(* IEC 61131-3 sources: daoli-st-library/DL_MathData (part 11) *)

(* ---- FC_DL_CubicBezierEval.st ---- *)
(*==============================================================================
 * 组件名称 (Component)  : FC_DL_CubicBezierEval
 * 所属子库 (Sublibrary) : DL_MathData
 * 当前版本 (Version)    : 1.0.0
 * 兼容性   (Platform)   : CODESYS 3.5+ / TwinCAT 3 / 汇川 InoProShop / 施耐德 Machine Expert
 *                         仅依赖 Standard.library 与 LREAL 四则运算，零厂商私有库
 * 功能描述 (Function)   : 一维标量三次贝塞尔曲线求值。给定四个控制点 P0~P3 与参数 t，
 *                         按 De Casteljau 递推（三级线性插值）求点值 fValue，并给出对 t 的
 *                         一阶导数 fTangent。选择 De Casteljau 而非多项式展开的理由：三次
 *                         Bernstein 展开在 t 接近 0/1 时会出现大系数相消（P0 与 P1 量级接近时
 *                         有效位丢失），De Casteljau 每级只做凸组合，数值稳定且中间量有界。
 * 分工声明 (Scope)      : 本件是**参数曲线求值**（已知控制点，求任意 t 处点与切线）；
 *                         `FC_DL_CubicSplineInterp` 是**数据点插值**（已知离散样本点，构造
 *                         分段三次样条后插值）。二者数学对象不同（Bernstein 基 vs 三次样条基），
 *                         不可互换调用：把本件当插值用会得到穿过控制包络的曲线而非过样本点曲线。
 * 接口     (Interface)  : 输入 fP0 / fP1 / fP2 / fP3 四个控制点标量值、fT 曲线参数（域 [0,1]，
 *                         越域钳制）；输出 fValue 点值、fTangent 一阶导数值、bClamped 参数
 *                         越域钳制标记、uErrorId 事件码；返回值 BOOL = TRUE 表示本次结果有效。
 * 边界     (Boundary)   : ① 参数越域（fT < 0 或 fT > 1）钳到端点并置 bClamped，不报错（钳制
 *                         是可预期的调用方行为，非故障）；
 *                         ② 任一输入非有限（NaN / ±Inf）→ 输出 0、置故障码、返回 FALSE，
 *                         绝不向下游传播 NaN（下游联锁会把 NaN 比较结果全判 FALSE 而静默失效）；
 *                         ③ 结果非有限复检兜底（防御纵深，正常域内不可能触发）；
 *                         ④ 纯函数零状态，无 TON / 边沿实例（R6 / R7 本件标注 N/A：无顺序状态机，
 *                         无实例调用，非法状态不可能出现）；
 *                         ⑤ 零全局耦合（无 GVL / 无物理地址）。
 * 判等例外 (Exception)  : 本件非有限判定使用 `x <> x`（NaN 自反）与 `(x-x) <> (x-x)`（Inf 差值
 *                         自减），此为**浮点判等禁令的唯一例外**（R79 / 机检 G6 白名单），
 *                         不得据此推断本件允许对量值使用 `=` / `<>`：量值比较在本件中不存在。
 * 码表     (Codes)      : 16#0001_03ED 故障级：贝塞尔求值故障（输入非有限 / 输出非有限复检失败），
 *                         本件单码，不细分（纯函数无归因成员，原因由入参侧唯一确定）。
 *                         16#0001_04B0 信息级：本次求值正常完成（供上层区分「未调用」与「调用成功」）。
 *                         加码反证（R90）：正常完成与「参数被钳制」在 fValue / fTangent 上不可区分
 *                         （钳制后 t 落到端点，结果与恰好传入端点值完全一致），故须以一码留痕；
 *                         钳制本身另有 bClamped 布尔出口，不再单立钳制码。
 *                         码段说明：0001 段故障子带 03xx / 信息子带 04xx，本件取 03ED / 04B0
 *                         （源码实扫该两槽为空，续接同子带已用最大值，未回填碎片孔洞）。
 * 开源溯源 (Origin)     : 道莅自研 clean-room（参考 Bernstein 基与 De Casteljau 公开算法定义，
 *                         零代码行复制；t2-1-lgf 数学子族）
 * 修订历史 (Revision)   : 2026-11-19  v1.0.0  R45 首版（批次 1 · 序号 4）
 *==============================================================================*)

FUNCTION FC_DL_CubicBezierEval : BOOL
VAR_INPUT
    fP0 : LREAL := 0.0;      // 控制点 P0 标量值（曲线起点），须有限 [工程单位] / Control point P0, curve start, must be finite
    fP1 : LREAL := 0.0;      // 控制点 P1 标量值（起点切线方向控制），须有限 [工程单位] / Control point P1, start tangent control
    fP2 : LREAL := 0.0;      // 控制点 P2 标量值（终点切线方向控制），须有限 [工程单位] / Control point P2, end tangent control
    fP3 : LREAL := 0.0;      // 控制点 P3 标量值（曲线终点），须有限 [工程单位] / Control point P3, curve end
    fT  : LREAL := 0.0;      // 曲线参数，有效域 0.0 ~ 1.0（越域钳制） [-] / Curve parameter, domain 0.0..1.0, out-of-range clamped
END_VAR
VAR_OUTPUT
    fValue   : LREAL;        // 曲线点值 B(t) [工程单位] / Curve point value B(t)
    fTangent : LREAL;        // 一阶导数 dB/dt（对 t 求导，非对弧长） [工程单位/参数] / First derivative dB/dt w.r.t. t
    bClamped : BOOL;         // 参数越域钳制标记 [-] / Parameter clamp flag
    uErrorId : UDINT;        // 事件码，0 = 无事件 / Event code, 0 = no event
END_VAR
VAR
    fTs      : LREAL;        // 钳制后的参数 t [-] / Clamped parameter t
    fOmT     : LREAL;        // 补参数 (1 - t) [-] / Complement parameter (1 - t)
    fQ0      : LREAL;        // 一级插值节点 Q0 [工程单位] / Level-1 node Q0
    fQ1      : LREAL;        // 一级插值节点 Q1 [工程单位] / Level-1 node Q1
    fQ2      : LREAL;        // 一级插值节点 Q2 [工程单位] / Level-1 node Q2
    fR0      : LREAL;        // 二级插值节点 R0 [工程单位] / Level-2 node R0
    fR1      : LREAL;        // 二级插值节点 R1 [工程单位] / Level-2 node R1
    fDiff01  : LREAL;        // 控制点差 P1 - P0 [工程单位] / Control point difference P1 - P0
    fDiff12  : LREAL;        // 控制点差 P2 - P1 [工程单位] / Control point difference P2 - P1
    fDiff23  : LREAL;        // 控制点差 P3 - P2 [工程单位] / Control point difference P3 - P2
    bNonFin  : BOOL;         // 输入非有限判定结果 [-] / Non-finite input verdict
END_VAR
VAR CONSTANT
    DL_BEZ_ORDER : LREAL := 3.0;   // 三次曲线阶数乘子（导数系数），编译期常量 [-] / Cubic order multiplier for derivative, compile-time constant
END_VAR

(* —— 段 1：返回值与输出预置（任何早退路径都不留脏值） —— *)
FC_DL_CubicBezierEval := FALSE;      // 返回值预置无效 / Preset return value invalid
fValue   := 0.0;                     // 点值预置 0，故障相即安全侧 / Point value preset 0, safe side in fault
fTangent := 0.0;                     // 切线预置 0 / Tangent preset 0
bClamped := FALSE;                   // 钳制标记预置 FALSE / Clamp flag preset FALSE
uErrorId := 16#0000_0000;            // 事件码预置无事件 / Event code preset none

(* —— 段 2：域闸（先判后算，禁算完再兜） —— *)
bNonFin := (fP0 <> fP0) OR (fP1 <> fP1) OR (fP2 <> fP2) OR (fP3 <> fP3) OR (fT <> fT)          // NaN 自反判（判等禁令唯一例外） / NaN self-reflexive test
        OR ((fP0 - fP0) <> (fP0 - fP0)) OR ((fP1 - fP1) <> (fP1 - fP1))                        // P1 差值自减判 Inf / Inf test on P1 via self-subtraction
        OR ((fP2 - fP2) <> (fP2 - fP2)) OR ((fP3 - fP3) <> (fP3 - fP3))                        // P2 / P3 差值自减判 Inf / Inf test on P2 and P3
        OR ((fT - fT) <> (fT - fT));                                                            // 参数差值自减判 Inf / Inf test on the parameter
IF bNonFin THEN
    uErrorId := 16#0001_03ED;        // 故障级：输入非有限，输出保持 0 / Fault-level: non-finite input, outputs stay zero
    RETURN;                          // 不抛异常，直接带码返回 / Return with code, no exception
END_IF

(* —— 段 3：参数钳制（越域钳到 [0,1] 并置标记） —— *)
IF fT < 0.0 THEN
    fTs := 0.0;                      // 下界钳制 / Clamp to lower bound
    bClamped := TRUE;                // 置钳制标记 / Set clamp flag
ELSIF fT > 1.0 THEN
    fTs := 1.0;                      // 上界钳制 / Clamp to upper bound
    bClamped := TRUE;                // 置钳制标记 / Set clamp flag
ELSE
    fTs := fT;                       // 域内直通 / Pass through inside domain
END_IF
fOmT := 1.0 - fTs;                   // 补参数 (1 - t) / Complement parameter

(* —— 段 4：De Casteljau 三级递推（委托内核，凸组合有界） —— *)
fQ0 := fOmT * fP0 + fTs * fP1;       // 一级插值 Q0 / Level-1 interpolation Q0
fQ1 := fOmT * fP1 + fTs * fP2;       // 一级插值 Q1 / Level-1 interpolation Q1
fQ2 := fOmT * fP2 + fTs * fP3;       // 一级插值 Q2 / Level-1 interpolation Q2
fR0 := fOmT * fQ0 + fTs * fQ1;       // 二级插值 R0 / Level-2 interpolation R0
fR1 := fOmT * fQ1 + fTs * fQ2;       // 二级插值 R1 / Level-2 interpolation R1
fValue := fOmT * fR0 + fTs * fR1;    // 三级插值 = 曲线点值 / Level-3 interpolation = curve point value
fDiff01 := fP1 - fP0;                // 起点段差 / Start segment difference
fDiff12 := fP2 - fP1;                // 中段差 / Middle segment difference
fDiff23 := fP3 - fP2;                // 终点段差 / End segment difference
fTangent := DL_BEZ_ORDER * ( fOmT * fOmT * fDiff01
                           + 2.0 * fOmT * fTs * fDiff12
                           + fTs * fTs * fDiff23 );   // Bernstein 导数式 dB/dt / Bernstein derivative dB/dt

(* —— 段 5：结果非有限复检兜底（防御纵深） —— *)
IF (fValue <> fValue) OR ((fValue - fValue) <> (fValue - fValue))
   OR (fTangent <> fTangent) OR ((fTangent - fTangent) <> (fTangent - fTangent)) THEN
    fValue   := 0.0;                 // 复检失败：点值归 0 / Recheck failed: point value zeroed
    fTangent := 0.0;                 // 复检失败：切线归 0 / Recheck failed: tangent zeroed
    uErrorId := 16#0001_03ED;        // 故障级：输出非有限 / Fault-level: non-finite output
    RETURN;                          // 带码返回 / Return with code
END_IF

(* —— 段 6：正常出口 —— *)
uErrorId := 16#0001_04B0;            // 信息级：求值正常完成 / Info-level: evaluation completed
FC_DL_CubicBezierEval := TRUE;       // 返回值置有效 / Return value valid

END_FUNCTION

(* ---- FC_DL_CubicSplineInterp.st ---- *)
(*
  FC_DL_CubicSplineInterp  —  自然三次样条插值与斜率输出 / Natural cubic spline interpolation with slope output
  分类 Category : DL_MathData
  码位 Code     : 16#05_0_01
  版本 Version  : 1.0.0
  来源标签 Tag  : t2-1-lgf-math
  溯源 Source   : LGF Math 语义借鉴 · clean-room 实现，仅借分类/参数域/命名，未复制源码行
  功能 Function : 1) 自然三次样条（二阶导三对角求解，Thomas 追赶法，WHILE 带死锁计数器上限 = 节点数 + 1）；
                  2) 同时输出插值值与一阶导数（斜率），供曲线跟踪/前馈使用；
                  3) 越界不外推：钳到端点并置 bInRange := FALSE。
  边界 Boundary : ① nPointCount < 2 判无效；
                  ② 节点 X 非严格递增（含相等）拒绝求值并置码，不做静默排序；
                  ③ fQueryX 越界 → 钳到端点、bInRange := FALSE、不外推；
                  ④ 三对角主元近零（|主元| < 1E-12）判节点病态置码；
                  ⑤ 节点数超 nMaxNode 组态上限拒绝（防静态数组越界）；
                  ⑥ 节点坐标非有限（NaN/Inf）拒绝求值（FB32-7 保持槽非有限闸）。
  依赖 Depends  : 无（纯 IEC 61131-3 标准运算，零库内内核可委托；SQRT/MOD 原语未使用）

  码表 Error codes（本件格 05_0_01，子码步进 +0x10）:
    16#0005_0501 故障级：组态非法（节点数 < 2 / 节点数超 nMaxNode / 节点 X 非严格递增 / 主元近零病态 / 节点非有限）
    16#0005_0511 信息级：查询点越界已钳到端点且不外推（不置 bError）

  修订历史 Revision :
    2026-11-18  v1.0.0  R36 首版入库（W1 窗次件）
*)

FUNCTION FC_DL_CubicSplineInterp : BOOL
VAR_INPUT
    afX        : ARRAY[0..63] OF LREAL;   // 节点横坐标表，要求严格递增 [任意工程单位] / Knot abscissa table, strictly increasing
    afY        : ARRAY[0..63] OF LREAL;   // 节点纵坐标表 [任意工程单位] / Knot ordinate table
    nPointCount : UINT := 0;              // 有效节点数 [个]，域 2 ~ nMaxNode / Effective knot count, domain 2..nMaxNode
    nMaxNode   : UINT := 64;              // 组态节点上限 [个]，域 2 ~ 64（静态数组上界保护）/ Configured max knot count
    fQueryX    : LREAL := 0.0;            // 查询横坐标 [任意工程单位] / Query abscissa
END_VAR
VAR_OUTPUT
    fOutY      : LREAL;                   // 插值结果 [任意工程单位]，无效时为 0 / Interpolated ordinate, 0 when invalid
    fOutSlope  : LREAL;                   // 一阶导数（斜率）[单位/单位]，无效时为 0 / First derivative, 0 when invalid
    bInRange   : BOOL;                    // 查询点是否落在节点区间内（FALSE 表示已钳到端点）/ Query inside knot span
    bValid     : BOOL;                    // 结果有效标志 / Result valid flag
    bError     : BOOL;                    // 故障标志，与故障级码配对 / Fault flag paired with fault code
    nErrId     : UDINT;                   // 事件码，0 = 无事件 / Event code, 0 = no event
END_VAR
VAR
    nCount     : INT;                                  // 生效节点数整型副本 [个] / Integer copy of knot count
    nLast      : INT;                                  // 末节点索引（nCount - 1）[1] / Last knot index
    i          : INT;                                  // 三对角求解行索引 [1] / Tridiagonal row index
    nGuard     : INT;                                  // 追赶快照死锁计数器 [1] / Back-substitution deadlock counter
    fHiPrev    : LREAL;                                // 左邻区间宽度 x[i]-x[i-1] [单位] / Left span width
    fHiNext    : LREAL;                                // 右邻区间宽度 x[i+1]-x[i] [单位] / Right span width
    fAlpha     : LREAL;                                // 追赶法右端项 [单位] / Thomas right-hand term
    fPivot     : LREAL;                                // 主元（对角元）[单位] / Pivot of tridiagonal system
    fQuery     : LREAL;                                // 生效查询横坐标（钳定后）[单位] / Effective (clamped) query abscissa
    fH         : LREAL;                                // 命中区间宽度 [单位] / Hit span width
    fA         : LREAL;                                // 左权 (x[i+1]-q)/h [1] / Left blend weight
    fB         : LREAL;                                // 右权 (q-x[i])/h [1] / Right blend weight
    nSeg       : INT;                                   // 命中区间左端索引 [1] / Hit span left index
    bFound     : BOOL;                                  // 区间查找命中标志 / Span found flag
    bMono      : BOOL;                                  // 节点严格递增检查标志 / Strict monotonic check flag
    bBad       : BOOL;                                  // 节点非有限标志 / Non-finite knot flag
    afM        : ARRAY[0..63] OF LREAL;                // 二阶导解向量 m[i] [单位] / Second derivative solution vector
    afL        : ARRAY[0..63] OF LREAL;                // 追赶法下对角 l[i] [单位] / Thomas lower diagonal
    afMu       : ARRAY[0..63] OF LREAL;                // 追赶法消元系数 mu[i] [1] / Thomas elimination coefficient
    afZ        : ARRAY[0..63] OF LREAL;                // 追赶法变换后右端 z[i] [单位] / Thomas transformed right-hand side
END_VAR
VAR CONSTANT
    DL_NODE_MIN : UINT  := 2;               // 节点数下限 [个]，单点无法定义斜率 / Minimum knot count
    DL_NODE_MAX : UINT  := 64;              // 节点数硬上限 [个]，等于数组上界 + 1 / Hard upper bound of knots
    DL_PIVOT_EPS : LREAL := 1.0E-12;       // 主元判零容差 [1]，低于此值判病态 / Pivot zero tolerance
    DL_EPS      : LREAL := 1.0E-12;        // 通用判零容差 [1] / Generic zero tolerance
END_VAR

(* —— 段 0：返回值与输出预置安全值 —— *)
FC_DL_CubicSplineInterp := FALSE;   // 返回布尔：FALSE = 本拍无有效结果
fOutY     := 0.0;                   // 插值结果预置 0
fOutSlope := 0.0;                   // 斜率预置 0
bInRange  := FALSE;                 // 区间内标志预置 FALSE
bValid    := FALSE;                 // 有效标志预置 FALSE
bError    := FALSE;                 // 故障标志预置 FALSE
nErrId    := 0;                     // 事件码预置 0
bFound    := FALSE;                 // 区间查找标志预置 FALSE
bMono     := TRUE;                  // 单调性假定成立
bBad      := FALSE;                 // 非有限假定不成立
nCount    := UINT_TO_INT(nPointCount);  // 节点数整型副本 [个]

(* —— 段 1：组态域闸（节点数与上限，先于任何数组访问） —— *)
IF (nCount < DL_NODE_MIN) OR (nCount > DL_NODE_MAX) THEN
    nErrId := 16#0005_0501;         // 故障级：节点数越 [2, 64] 域
    bError := TRUE;                 // 故障标志置位（R45 配对）
    RETURN;                         // 域闸命中不求值
END_IF
IF (nMaxNode < DL_NODE_MIN) OR (nMaxNode > DL_NODE_MAX) THEN
    nErrId := 16#0005_0501;         // 故障级：组态上限越域
    bError := TRUE;                 // 故障标志置位（R45 配对）
    RETURN;                         // 域闸命中不求值
END_IF
IF nPointCount > nMaxNode THEN
    nErrId := 16#0005_0501;         // 故障级：实际节点数超组态上限（防越界，不静默截断）
    bError := TRUE;                 // 故障标志置位（R45 配对）
    RETURN;                         // 域闸命中不求值
END_IF
IF (fQueryX <> fQueryX) OR ((fQueryX - fQueryX) <> (fQueryX - fQueryX)) THEN
    nErrId := 16#0005_0501;         // 故障级：查询横坐标非有限
    bError := TRUE;                 // 故障标志置位（R45 配对）
    RETURN;                         // 域闸命中不求值
END_IF
nLast := nCount - 1;                // 末节点索引 [1]

(* —— 段 2：节点表体检（严格递增 + 非有限），任一不满足拒绝求值 —— *)
FOR i := 0 TO nLast DO
    IF (afX[i] <> afX[i]) OR ((afX[i] - afX[i]) <> (afX[i] - afX[i])) THEN
        bBad := TRUE;               // 节点横坐标非有限
    END_IF
    IF (afY[i] <> afY[i]) OR ((afY[i] - afY[i]) <> (afY[i] - afY[i])) THEN
        bBad := TRUE;               // 节点纵坐标非有限
    END_IF
END_FOR
IF bBad THEN
    nErrId := 16#0005_0501;         // 故障级：节点表含非有限值
    bError := TRUE;                 // 故障标志置位（R45 配对）
    RETURN;                         // 不求值
END_IF
FOR i := 1 TO nLast DO
    IF afX[i] - afX[i - 1] <= 0.0 THEN
        bMono := FALSE;             // 非严格递增（含相等与倒序）
    END_IF
END_FOR
IF NOT bMono THEN
    nErrId := 16#0005_0501;         // 故障级：节点 X 非严格递增，拒绝求值（不做静默排序）
    bError := TRUE;                 // 故障标志置位（R45 配对）
    RETURN;                         // 不求值
END_IF

(* —— 段 3：自然样条二阶导求解（Thomas 追赶法，主元近零判病态） —— *)
afM[0] := 0.0;                      // 自然边界：首端二阶导为 0
afM[nLast] := 0.0;                  // 自然边界：末端二阶导为 0
afL[0] := 1.0;                      // 追赶法初值
afMu[0] := 0.0;                     // 追赶法初值
afZ[0] := 0.0;                      // 追赶法初值
FOR i := 1 TO (nLast - 1) DO
    fHiPrev := afX[i] - afX[i - 1];                                  // 左邻区间宽度 [单位]
    fHiNext := afX[i + 1] - afX[i];                                  // 右邻区间宽度 [单位]，递增性已证明 > 0
    fAlpha := 3.0 / fHiNext * (afY[i + 1] - afY[i]) - 3.0 / fHiPrev * (afY[i] - afY[i - 1]);  // 右端项
    fPivot := 2.0 * (afX[i + 1] - afX[i - 1]) - fHiPrev * afMu[i - 1];                        // 主元
    IF ABS(fPivot) < DL_PIVOT_EPS THEN
        nErrId := 16#0005_0501;     // 故障级：三对角主元近零，节点病态
        bError := TRUE;             // 故障标志置位（R45 配对）
        RETURN;                     // 不出结论
    END_IF
    afL[i] := fPivot;                                               // 保存消元主元
    afMu[i] := fHiNext / afL[i];                                    // 消元系数（主元已证明非零）
    afZ[i] := (fAlpha - fHiPrev * afZ[i - 1]) / afL[i];             // 变换后右端
END_FOR
afM[nLast] := 0.0;                  // 自然边界复核（末端）
nGuard := 0;                        // 死锁计数器清零
i := nLast - 1;                     // 回代起点
WHILE (i >= 1) AND (nGuard <= (nCount + 1)) DO
    afM[i] := afZ[i] - afMu[i] * afM[i + 1];                        // 回代求二阶导
    i := i - 1;                                                     // 索引递减
    nGuard := nGuard + 1;                                           // 死锁计数器自增
END_WHILE
IF nGuard > (nCount + 1) THEN
    nErrId := 16#0005_0501;         // 故障级：回代未在节点数 + 1 步内收敛（结构性防御）
    bError := TRUE;                 // 故障标志置位（R45 配对）
    RETURN;                         // 不出结论
END_IF

(* —— 段 4：定位命中区间（线性查找，不外推：越界钳到端点） —— *)
fQuery := fQueryX;                  // 生效查询横坐标初值
IF fQueryX < afX[0] THEN
    fQuery := afX[0];               // 左越界钳到首端，不外推
    bInRange := FALSE;              // 标记越界
ELSIF fQueryX > afX[nLast] THEN
    fQuery := afX[nLast];           // 右越界钳到末端，不外推
    bInRange := FALSE;              // 标记越界
ELSE
    bInRange := TRUE;               // 落在节点区间内
END_IF
nSeg := 0;                          // 区间左端索引初值
FOR i := 0 TO (nLast - 1) DO
    IF (fQuery >= afX[i]) AND (fQuery <= afX[i + 1]) THEN
        nSeg := i;                  // 命中区间 [x[i], x[i+1]]
        bFound := TRUE;             // 查找命中
        EXIT;                       // 唯一区间（严格递增保证）
    END_IF
END_FOR
IF NOT bFound THEN
    nSeg := nLast - 1;              // 端点等值数值落空的兜底：取末区间
END_IF

(* —— 段 5：区间内求值与斜率（h 已证明 > 0，无除零风险） —— *)
fH := afX[nSeg + 1] - afX[nSeg];                                        // 命中区间宽度 [单位]
IF fH <= 0.0 THEN
    nErrId := 16#0005_0501;         // 故障级：命中区间宽度非正（数值退化）
    bError := TRUE;                 // 故障标志置位（R45 配对）
    RETURN;                         // 不出结论
END_IF
fA := (afX[nSeg + 1] - fQuery) / fH;                                    // 左权 [1]
fB := (fQuery - afX[nSeg]) / fH;                                        // 右权 [1]
fOutY := fA * afY[nSeg] + fB * afY[nSeg + 1]
       + ((fA * fA * fA - fA) * afM[nSeg] + (fB * fB * fB - fB) * afM[nSeg + 1]) * fH * fH / 6.0;  // 插值结果
fOutSlope := (afY[nSeg + 1] - afY[nSeg]) / fH
           - (3.0 * fA * fA - 1.0) / 6.0 * fH * afM[nSeg]
           + (3.0 * fB * fB - 1.0) / 6.0 * fH * afM[nSeg + 1];           // 一阶导数

(* —— 段 6：结果非有限复检 + 越界信息码 + 有效标志 —— *)
IF (fOutY <> fOutY) OR ((fOutY - fOutY) <> (fOutY - fOutY)) THEN
    fOutY := 0.0;                   // 非有限复检兜底
    fOutSlope := 0.0;               // 斜率同步兜底
    nErrId := 16#0005_0501;         // 故障级：插值结果非有限
    bError := TRUE;                 // 故障标志置位（R45 配对）
    RETURN;                         // 不出结论
END_IF
IF NOT bInRange THEN
    nErrId := 16#0005_0511;         // 信息级：查询点越界已钳到端点（信息级不置 bError）
END_IF
bValid := TRUE;                     // 结果有效（越界钳定亦有效，但 bInRange 已置 FALSE 提示）
FC_DL_CubicSplineInterp := TRUE;    // 返回布尔：TRUE = 本拍有可交付结果

END_FUNCTION

(* ---- FC_DL_CvdFilmStressCalc.st ---- *)
(*
  DL Factory R88 | FC_DL_CvdFilmStressCalc
  功能：Stoney 式算薄膜应力 σ=E_s·t_s²/(6(1-ν)·t_f·R)，曲率半径取绝对值、符号由曲率方向给定，超 300 MPa 提示
  开源溯源：无（clean-room 自研，依据公开工艺公式 Stoney 薄膜应力式，许可证=MIT，借鉴点=公式结构）
  规则：R1-R16 全遵守；R88 简单件标量形（纯标量入参出参，无循环体、无方法、无属性、无数组）
*)
FUNCTION FC_DL_CvdFilmStressCalc : REAL
VAR_INPUT
    fSubstModulusGPa : REAL := 200.0; // 基片双轴模量 E_s（Si(100) 约 180 GPa） [GPa] / substrate biaxial modulus [GPa]
    fSubstThkUm : REAL := 725.0; // 基片厚度 t_s [µm] / substrate thickness [um]
    fPoissonNu : REAL := 0.28; // 基片泊松比 ν（Si 约 0.28） [-] / Poisson ratio [-]
    fFilmThkUm : REAL := 1.0; // 薄膜厚度 t_f（须远小于 t_s） [µm] / film thickness [um]
    fCurvRadiusM : REAL := 10.0; // 曲率半径 R（带符号：正=上凸/张应力，负=下凹/压应力） [m] / signed radius [m]
    fLimitMPa : REAL := 300.0; // 应力绝对值报警上限 [MPa] / absolute stress alarm limit [MPa]
END_VAR
VAR_OUTPUT
    fStressMPa : REAL; // 薄膜应力 σ（正=张应力，负=压应力） [MPa] / film stress, positive is tensile [MPa]
    xOverLimit : BOOL; // TRUE=应力绝对值超过上限 [-] / TRUE when the absolute value is above the limit [-]
END_VAR
VAR
    fTsM : REAL; // 基片厚度换算为 m [m] / substrate thickness in metres [m]
    fTfM : REAL; // 薄膜厚度换算为 m（除零判据） [m] / film thickness in metres, the divisor [m]
    fDenom : REAL; // 分母 6(1-ν)·t_f·R_abs（除零判据） [m²] / denominator, the divisor [m^2]
    fMagMPa : REAL; // 应力幅值（未加符号） [MPa] / stress magnitude [MPa]
END_VAR

// 段 1｜出口预置
FC_DL_CvdFilmStressCalc := -1.0; // 哨兵返回 -1（无效） [-] / sentinel return -1, invalid [-]
fStressMPa := 0.0; // 应力预置零 [MPa] / stress preset zero [MPa]
xOverLimit := FALSE; // 超限位预置 FALSE（未判定前不报警） [-] / over-limit flag preset false [-]

// 段 2｜非有限拦截 + 域闸
IF NOT (fSubstModulusGPa > -1.0E30 AND fSubstModulusGPa < 1.0E30) OR NOT (fSubstThkUm > -1.0E30 AND fSubstThkUm < 1.0E30) OR NOT (fPoissonNu > -1.0E30 AND fPoissonNu < 1.0E30) THEN
    RETURN; // 模量/基片厚/泊松比任一非有限即拒算 [-] / any non finite input rejected [-]
END_IF
IF NOT (fFilmThkUm > -1.0E30 AND fFilmThkUm < 1.0E30) OR NOT (fCurvRadiusM > -1.0E30 AND fCurvRadiusM < 1.0E30) OR NOT (fLimitMPa > -1.0E30 AND fLimitMPa < 1.0E30) THEN
    RETURN; // 膜厚/曲率半径/上限任一非有限则判据静默失效，故先拦 [-] / these pins must be finite [-]
END_IF
IF fSubstModulusGPa <= 0.0 OR fSubstThkUm < 1.0E-9 OR fFilmThkUm < 1.0E-9 THEN
    RETURN; // 模量正域闸 + 厚度正域闸（分母因子不得为零） [GPa, µm] / positive modulus and thicknesses
END_IF
IF fPoissonNu <= -1.0 OR fPoissonNu >= 0.5 OR ABS(fCurvRadiusM) < 1.0E-9 OR fLimitMPa <= 0.0 THEN
    RETURN; // 泊松比开区间闸 (-1,0.5) + 曲率绝对值闸 + 上限正域闸 [-] / Poisson, radius and limit gates
END_IF

// 段 3｜计算（Stoney 式，长度统一换算到 m、模量换算到 Pa，末步转 MPa）
fTsM := fSubstThkUm * 1.0E-6; // µm × 1e-6 m/µm = m，基片厚换算 [m] / [um] x [m/um] = [m]
fTfM := fFilmThkUm * 1.0E-6; // µm × 1e-6 m/µm = m，膜厚换算 [m] / [um] x [m/um] = [m]
fDenom := 6.0 * (1.0 - fPoissonNu) * fTfM * ABS(fCurvRadiusM); // 无量纲 × 无量纲 × m × m = m²，分母 [m²] / [m^2]
IF fDenom < 1.0E-9 THEN
    RETURN; // 除法前分母闸：6(1-ν)t_f·R 必须大于 1E-9 才可作除数 [m²] / denominator gate [m^2]
END_IF
fMagMPa := fSubstModulusGPa * 1.0E9 * fTsM * fTsM / fDenom * 1.0E-6; // Pa × m² ÷ m² = Pa，再 ×1e-6 转 MPa [MPa] / [MPa]
IF fCurvRadiusM < 0.0 THEN
    fStressMPa := -fMagMPa; // 负曲率对应压应力（符号约定），幅值来自上式的绝对半径 [MPa] / compressive [MPa]
ELSE
    fStressMPa := fMagMPa; // 正曲率对应张应力（符号约定），幅值来自上式的绝对半径 [MPa] / tensile [MPa]
END_IF

// 段 4｜判定与饱和
IF NOT (fStressMPa > -1.0E30 AND fStressMPa < 1.0E30) THEN
    RETURN; // 结果非有限再拦一次（防溢出成 Inf） [MPa] / re-check the result for finiteness [MPa]
END_IF
xOverLimit := ABS(fStressMPa) > fLimitMPa; // 按绝对值与上限直比（张压同判） [MPa] / compare the magnitude [MPa]

// 段 5｜出口自检
IF fTfM >= fTsM THEN RETURN; END_IF // 出口自检：Stoney 式前提是薄膜远薄于基片，t_f>=t_s 时结果不可信 [m] / premiss violated
FC_DL_CvdFilmStressCalc := fStressMPa; // 返回薄膜应力（正=张，负=压） [MPa] / return the film stress [MPa]
END_FUNCTION

(* ---- FC_DL_DateAddDays.st ---- *)
(*
    FC_DL_DateAddDays —— DATE 加天数偏移
    ------------------------------------------------------------------
    分类      : DL_MathData / TimeArith
    前缀      : FC_DL_
    版本      : 1.0.0
    溯源      : IEC 61131-3 标准语义的道莅防御性实现（日期 + 天数 → 日期，可负偏移）；
                经天数路径委托平台内建 DATE_TO_DINT / DINT_TO_DATE 完成历法换算，
                本件不重实现历法内核；
                偏移钳位、溢出预判、双出口错误分级与码位 100% 自有；
                clean-room 重写，未复制任何闭源厂商源码，参考实现仅限 MIT/Apache 许可
    平台      : 纯 IEC 61131-3，CODESYS V3.5+ / TwinCAT 3 / InoProShop 通用
    作者      : 道莅代码库 · PLC编程专家（R20）
    ------------------------------------------------------------------
    功能说明  : 保质期到日子、交期推算、下次保养日（今天 + 90 天）、点检周期回推（今天 − 30 天）
                这类现场每天都在用的算术。日历加法不能靠秒数硬加：夏令时与闰秒都不参与
                工业日期的语义，天数路径才是唯一稳定口径。
                核心防御：① 统一走天数路径（先 DATE_TO_DINT，加偏移后再 DINT_TO_DATE），
                   不做 DT 秒级加减——秒级加减在跨闰日的边界上会差一天，而这一天
                   对保质期判定的意义不用解释；
                ② 溢出用减法比较预判，不用加法后回查符号位：nWork > 上限 − nBase
                   这类判据在任何整数表示下都成立，禁「先加再判是否变号」的写法
                   （带符号溢出的回绕行为在平台上并不一定有保证）；
                ③ 偏移超 ±36500 天（±100 年）先钳位并发信息级：排程里出现 ±100 年
                   必然是单位错（毫秒当秒填），钳位后可算但不静默；
                ④ 结果早于纪元或超容器域一律返回纪元日并置 bValid = FALSE，不做饱和——
                   饱和会伪造日期（把越界算成 1970-01-01），台账上看不出异常；
                ⑤ 天数上界与 FC_DL_DateToDintDays / FC_DL_DintDaysToDate 用同一常量口径，
                   三件之间不会错位。
                职责边界：日期差值归 FC_DL_DateDiffDays；闰年原子归 FC_DL_LeapYearChk；
                纯天数双向转换归 FC_DL_DateToDintDays / FC_DL_DintDaysToDate。
    编译门槛  : 主路径依赖平台内建 DATE_TO_DINT / DINT_TO_DATE（天数口径），
                三平台标准库均提供。天数口径的平台差异见 FC_DL_DateToDintDays 的
                编译门槛段与 DL_DATE_DAYS_MAX 的保守取值；若实测口径不同只调该常量，
                本件的闸门顺序与出口不变。
    错误码    : 16#0001_042A 偏移超 ±36500 天（±100 年）已钳位——信息级，值可用但偏移已被限幅
                16#0001_042B 预留禁用（信息级，不得挪用）
                16#0001_035D 结果早于纪元——故障级，返回纪元日
                16#0001_035E 结果超 DATE 容器域——故障级，返回纪元日，不做饱和
                16#0001_035F 预留禁用（故障级，不得挪用）
    码位总账  : 16#0001_042A 用 / 16#0001_042B 预留 ｜ 16#0001_035D 用 / 16#0001_035E 用 / 16#0001_035F 预留
    状态机    : R6 标注 N/A —— 本组件为纯函数无顺序状态机，无 CASE 可写，非法状态不可能出现
    采样约定  : 本件无定时器、无沿检测、无状态；单拍纯计算，结论与任务周期无关。
    修订记录  : 2026-11-16 v1.0.0 首次入库（R20）
*)
FUNCTION FC_DL_DateAddDays : DATE
VAR_INPUT
    dateIn           : DATE;                  // 基准日期 [日期]，有效域 1970-01-01 起 / base date [date], domain starts at 1970-01-01
    nDays            : DINT;                  // 天数偏移，可负 [日]，有效域 −36500~36500 / day offset, signed [day], valid domain −36500 to 36500
END_VAR
VAR_OUTPUT
    eErr             : UDINT;                 // 错误码，0=正常 / error id, 0=ok
    bError           : BOOL;                  // 故障标志，eErr 为故障级时 TRUE / error flag, TRUE on fault-level eErr
    bValid           : BOOL;                  // 返回值是否可用（故障级为 FALSE）/ return usable, FALSE on fault level
    bClamped         : BOOL;                  // 偏移超 ±36500 天已钳位 / the offset was clamped into the span limit
END_VAR
VAR CONSTANT
    DL_DAYS_SPAN_MAX : DINT := 36500;         // 正向偏移钳位，约 ±100 年 [日] / forward offset clamp, about one hundred years [day]
    DL_DAYS_SPAN_NEG_MAX : DINT := -36500;    // 负向偏移钳位 [日] / backward offset clamp [day]
    DL_DATE_DAYS_MIN : DINT := 0;             // 纪元日，天数下界 [日] / the epoch day, lower bound [day]
    DL_DATE_DAYS_MAX : DINT := 65535;         // 保守容器口径上限，无符号 16 位天数顶 [日] / conservative container top [day]
    DL_EPOCH_DATE_ZERO : DATE := DATE#1970-01-01; // 纪元起始日期，故障缺省返回 / the epoch date returned on faults
END_VAR
VAR
    nBase            : DINT;                  // 基准日期天数中间量 [日] / base date in days since the epoch [day]
    nWork            : DINT;                  // 偏移副本，钳位后参与加法 [日] / offset copy, used after the clamp [day]
    nOut             : DINT;                  // 结果天数中间量 [日] / result day count intermediate [day]
    nLimit           : DINT;                  // 可用余量的减法判据中间量 [日] / headroom intermediate used by the subtraction test [day]
END_VAR

// 段 1｜返回值与错误状态预置 / segment 1, preset return value and error status
FC_DL_DateAddDays := DL_EPOCH_DATE_ZERO;      // 故障缺省返回纪元日 / fault default returns the epoch date
eErr := 0;                                    // 预置无错误 / preset no error
bError := FALSE;                              // 预置无故障 / preset no fault
bValid := FALSE;                              // 预置不可用，通过闸门后置位 / preset invalid, set TRUE after the gates
bClamped := FALSE;                            // 预置未钳位 / preset no clamp
nWork := nDays;                               // 取入参副本，绝不改动调用方数据 / copy the input, never modifies caller data
nOut := DL_DATE_DAYS_MIN;                     // 结果中间量清零 / clear the result intermediate

// 段 2｜偏移跨度量闸：超 ±100 年先钳位并如实登记（信息级）/ segment 2, span gate with an explicit info-level clamp
IF nWork > DL_DAYS_SPAN_MAX THEN
    nWork := DL_DAYS_SPAN_MAX;                // 正向钳位至 +36500 天 [日] / clamp to plus 36500 days [day]
    bClamped := TRUE;                         // 标记已钳位 / flag the clamp
    eErr := 16#0001_042A;                     // 信息级：偏移超跨度已钳位 / info level, the offset was clamped
ELSIF nWork < DL_DAYS_SPAN_NEG_MAX THEN
    nWork := DL_DAYS_SPAN_NEG_MAX;            // 负向钳位至 −36500 天 [日] / clamp to minus 36500 days [day]
    bClamped := TRUE;                         // 标记已钳位 / flag the clamp
    eErr := 16#0001_042A;                     // 信息级：偏移超跨度已钳位 / info level, the offset was clamped
END_IF

// 段 3｜基准日期域闸：基准本身必须在容器域内 / segment 3, base date domain gate
nBase := DATE_TO_DINT(dateIn);                // 日期 → 自纪元天数 [日] / date to days since the epoch [day]
IF nBase < DL_DATE_DAYS_MIN THEN
    eErr := 16#0001_035D;                     // 故障级：基准日期早于纪元 / fault level, the base date precedes the epoch
    bError := TRUE;                           // 置故障标志 / raise the error flag
    bValid := FALSE;                          // 返回值不可用 / flag the return as unusable
    FC_DL_DateAddDays := DL_EPOCH_DATE_ZERO;  // 确定缺省值：纪元日 / deterministic default of the epoch date
    RETURN;                                   // 出口 / exit
END_IF
IF nBase > DL_DATE_DAYS_MAX THEN
    eErr := 16#0001_035E;                     // 故障级：基准日期超容器域 / fault level, the base date exceeds the container
    bError := TRUE;                           // 置故障标志 / raise the error flag
    bValid := FALSE;                          // 返回值不可用 / flag the return as unusable
    FC_DL_DateAddDays := DL_EPOCH_DATE_ZERO;  // 确定缺省值：纪元日 / deterministic default of the epoch date
    RETURN;                                   // 出口 / exit
END_IF

// 段 4｜正向溢出预判：用「上限 − 基准」做减法比较，禁先加后判变号 / segment 4, forward overflow test by subtraction
IF nWork > DL_DATE_DAYS_MIN THEN
    nLimit := DL_DATE_DAYS_MAX - nBase;       // 剩余可用天数 [日] / remaining room in days [day]
    IF nWork > nLimit THEN
        eErr := 16#0001_035E;                 // 故障级：结果将超 DATE 容器域 / fault level, the result would exceed the container
        bError := TRUE;                       // 置故障标志 / raise the error flag
        bValid := FALSE;                      // 返回值不可用 / flag the return as unusable
        FC_DL_DateAddDays := DL_EPOCH_DATE_ZERO; // 确定缺省值：纪元日，不伪造日期 / deterministic default, no fabricated date
        RETURN;                               // 出口 / exit
    END_IF
ELSIF nWork < DL_DATE_DAYS_MIN THEN
    // 段 5｜负向溢出预判：可用余额同为负数，比较方向不变 / segment 5, backward overflow test
    nLimit := DL_DATE_DAYS_MIN - nBase;       // 负向可用余额，负值 [日] / backward headroom, a negative value [day]
    IF nWork < nLimit THEN
        eErr := 16#0001_035D;                 // 故障级：结果将早于纪元 / fault level, the result would precede the epoch
        bError := TRUE;                       // 置故障标志 / raise the error flag
        bValid := FALSE;                      // 返回值不可用 / flag the return as unusable
        FC_DL_DateAddDays := DL_EPOCH_DATE_ZERO; // 确定缺省值：纪元日 / deterministic default of the epoch date
        RETURN;                               // 出口 / exit
    END_IF
END_IF

// 段 6｜主体：溢出已排除，加法与内建还原均安全 / segment 6, the addition and the built-in are safe after the gates
nOut := nBase + nWork;                        // 结果天数 [日] / result day count [day]
FC_DL_DateAddDays := DINT_TO_DATE(nOut);      // 天数 → 日期 / days back to a date

// 段 7｜发布结果 / segment 7, publish the result
bValid := TRUE;                               // 域内结果可用 / the in-domain result is usable
bError := FALSE;                              // 信息级不置故障（双保险）/ info level never raises a fault, second line of defence
END_FUNCTION

(* ---- FC_DL_DateDiffDays.st ---- *)
(*
    FC_DL_DateDiffDays —— 两 DATE 之差天数（可负）
    ------------------------------------------------------------------
    分类      : DL_MathData / TimeArith
    前缀      : FC_DL_
    版本      : 1.0.0
    溯源      : IEC 61131-3 标准语义的道莅防御性实现（两个日期之间的天数差，可负）；
                经天数路径委托平台内建 DATE_TO_DINT 完成历法换算，本件不重实现历法内核；
                负值口径、方向标志、错误分级与码位 100% 自有；
                clean-room 重写，未复制任何闭源厂商源码，参考实现仅限 MIT/Apache 许可
    平台      : 纯 IEC 61131-3，CODESYS V3.5+ / TwinCAT 3 / InoProShop 通用
    作者      : 道莅代码库 · PLC编程专家（R20）
    ------------------------------------------------------------------
    功能说明  : 保质期余量、超期天数、保养逾期天数的判定原子：给两个日期，输出「从前者到后者
                过了多少天」，后者早于前者即为负。与 FC_DL_DateAddDays 构成判定原子对。
                核心防御：① 差值一律在 DINT 域内做：两个 DATE 都在容器域内，天数差模长必小于
                   65536，DINT 承载结构性不溢出——此论证是本件不设故障出口的依据；
                ② 负值是合法业务输出（超期天数就是负的余量），绝不钳到 0、绝不用绝对值：
                   把「已超期 3 天」抹平成「今天到期」是保质期逻辑最典型的静默错；
                ③ bNegative 单独回告方向，HMI 不必自己再比一次大小；
                ④ 本件五槽中信息 1 槽使用、故障 3 槽按规格预留——域外输入在类型域上
                   不可表达（DATE 值域由类型系统保证），故不虚构不存在的故障码。
                职责边界：日期加偏移归 FC_DL_DateAddDays；日期天数化归 FC_DL_DateToDintDays；
                本件只管两日期之间的差值。
    编译门槛  : 主路径依赖平台内建 DATE_TO_DINT（天数口径），三平台标准库均提供。
                若某平台 DATE 以秒承载，则差值单位为秒而非天——此差异由 DL_DATE_DAYS_MAX
                的实测锚定统一裁定（与 FC_DL_DateToDintDays 同源），本件闸门不受影响。
    错误码    : 16#0001_042C 差值为负（dateTo 早于 dateFrom），已如实输出——信息级，值可用
                16#0001_042D 预留禁用（信息级，不得挪用）
                16#0001_0360 预留（故障级，不得挪用）
                16#0001_0361 预留禁用（故障级，不得挪用）
                16#0001_0362 预留禁用（故障级，不得挪用）
    码位总账  : 16#0001_042C 用 / 16#0001_042D 预留 ｜ 16#0001_0360 预留 / 16#0001_0361 预留 / 16#0001_0362 预留
    状态机    : R6 标注 N/A —— 本组件为纯函数无顺序状态机，无 CASE 可写，非法状态不可能出现
    采样约定  : 本件无定时器、无沿检测、无状态；单拍纯计算，结论与任务周期无关。
    修订记录  : 2026-11-16 v1.0.0 首次入库（R20）
*)
FUNCTION FC_DL_DateDiffDays : DINT
VAR_INPUT
    dateFrom         : DATE;                  // 区间起始日期 [日期] / start date of the interval [date]
    dateTo           : DATE;                  // 区间结束日期 [日期]，早于起点即差值为负 / end date of the interval [date], earlier than the start yields a negative difference
END_VAR
VAR_OUTPUT
    eErr             : UDINT;                 // 错误码，0=正常 / error id, 0=ok
    bError           : BOOL;                  // 故障标志，本件无故障级出口，恒为 FALSE / error flag, always FALSE here as no fault exit exists
    bValid           : BOOL;                  // 返回值是否可用（本件恒为 TRUE）/ return usable, always TRUE here
    bNegative        : BOOL;                  // 差值为负（dateTo 早于 dateFrom）/ the difference is negative
END_VAR
VAR CONSTANT
    DL_DINT_ZERO     : DINT := 0;             // 有符号零常量，避免裸字面量 [日] / signed zero constant [day]
END_VAR
VAR
    nFrom            : DINT;                  // 起始日期天数 [日] / start date in days [day]
    nTo              : DINT;                  // 结束日期天数 [日] / end date in days [day]
    nDiff            : DINT;                  // 差值中间量，可负 [日] / difference intermediate, possibly negative [day]
END_VAR

// 段 1｜返回值与错误状态预置 / segment 1, preset return value and error status
FC_DL_DateDiffDays := DL_DINT_ZERO;           // 缺省返回 0 天 [日] / default returns zero days [day]
eErr := 0;                                    // 预置无错误 / preset no error
bError := FALSE;                              // 本件无故障级出口，恒 FALSE / no fault exit exists, always FALSE
bValid := FALSE;                              // 预置不可用，末段置位 / preset invalid, set TRUE in the last stage
bNegative := FALSE;                           // 预置非负差 / preset a non-negative difference
nDiff := DL_DINT_ZERO;                        // 中间量清零 / clear the intermediate

// 段 2｜取值：两日期各做一次显式标准转换 / segment 2, both dates are converted explicitly
nFrom := DATE_TO_DINT(dateFrom);              // 起始日期天数 [日] / start date in days [day]
nTo := DATE_TO_DINT(dateTo);                  // 结束日期天数 [日] / end date in days [day]

// 段 3｜求差：模长必小于 65536，DINT 承载结构性不溢出 / segment 3, the difference cannot overflow DINT
nDiff := nTo - nFrom;                         // 有符号天数差 [日] / signed difference in days [day]

// 段 4｜负值如实输出（超期余量语义，绝不抹平）/ segment 4, negative values are published as they are
IF nDiff < DL_DINT_ZERO THEN
    bNegative := TRUE;                        // 标记差值为负 / flag the negative difference
    eErr := 16#0001_042C;                     // 信息级：差值为负，已如实输出 / info level, a negative difference was published as is
END_IF

// 段 5｜发布结果 / segment 5, publish the result
FC_DL_DateDiffDays := nDiff;                  // 输出天数差 [日] / publish the difference in days [day]
bValid := TRUE;                               // 正负差值均为合法业务输出 / both signs are legal business results
bError := FALSE;                              // 信息级不置故障（双保险）/ info level never raises a fault, second line of defence
END_FUNCTION

(* ---- FC_DL_DateToDintDays.st ---- *)
(*
    FC_DL_DateToDintDays —— DATE 到自纪元起的天数
    ------------------------------------------------------------------
    分类      : DL_MathData / Convert
    前缀      : FC_DL_
    版本      : 1.0.0
    溯源      : IEC 61131-3 标准语义的道莅防御性实现（DATE → 自 1970-01-01 起天数）；
                委托平台内建 DATE_TO_DINT 完成天数口径换算，本件不重实现历法内核；
                纪元域闸门、保守容器口径钳位、错误分级与码位 100% 自有；
                clean-room 重写，未复制任何闭源厂商源码，参考实现仅限 MIT/Apache 许可
    平台      : 纯 IEC 61131-3，CODESYS V3.5+ / TwinCAT 3 / InoProShop 通用
    作者      : 道莅代码库 · PLC编程专家（R20）
    ------------------------------------------------------------------
    功能说明  : 把日历日期折成「自 1970-01-01 起的天数」整数，供保质期、台账天数化、
                保养周期差值与数据库整型列落库使用（日期型直接落库在各家平台的位型不一致）。
                核心防御：① 早于纪元的日期在调用内建前拦下，域外调用内建可得回绕大数；
                ② 天数超保守容器口径时按容器顶钳位并发信息级，值仍可用但已注明钳位——
                   钳位事件必须可被 HMI 看见，静默钳位是本件最易漏的缺陷；
                ③ 内建返回负天数视为容器溢出（与段 2 的域门同源但不同层），单独占故障码，
                   便于区分「组态给了 1970 前日期」与「平台 DATE 位型承载异常」两类根因。
                职责边界：天数还原归 FC_DL_DintDaysToDate；带偏移的日期推算归
                FC_DL_DateAddDays；日期差值归 FC_DL_DateDiffDays。
    编译门槛  : 主路径依赖平台内建 DATE_TO_DINT（天数口径）。三平台标准库均提供该内建，
                但天数口径本身的数值锚定存在平台差异：某些平台 DATE 以秒承载、部分以天承载。
                故 DL_DATE_DAYS_MAX 取 65535（无符号 16 位天数容器上限）的保守口径，
                编码前按目标平台实测锚定；若实测口径不同，仅调本常量，闸门与出口不动。
    错误码    : 16#0001_0410 天数超保守容器口径（65535），已按容器顶钳位——信息级，值仍可用但已钳位
                16#0001_0411 预留禁用（信息级，不得挪用）
                16#0001_0336 输入日期早于纪元（1970-01-01 之前）——故障级，返回 0
                16#0001_0337 DATE 输入非法或容器溢出（内建返回负天数）——故障级，返回 0
                16#0001_0338 预留禁用（故障级，不得挪用）
    码位总账  : 16#0001_0410 用 / 16#0001_0411 预留 ｜ 16#0001_0336 用 / 16#0001_0337 用 / 16#0001_0338 预留
    状态机    : R6 标注 N/A —— 本组件为纯函数无顺序状态机，无 CASE 可写，非法状态不可能出现
    采样约定  : 本件无定时器、无沿检测、无状态；单拍纯计算，结论与任务周期无关。
    修订记录  : 2026-11-16 v1.0.0 首次入库（R20）
*)
FUNCTION FC_DL_DateToDintDays : DINT
VAR_INPUT
    dateIn           : DATE;                  // 输入日期 [日期]，有效域 1970-01-01 起 / input date [date], domain starts at 1970-01-01
END_VAR
VAR_OUTPUT
    eErr             : UDINT;                 // 错误码，0=正常 / error id, 0=ok
    bError           : BOOL;                  // 故障标志，eErr 为故障级时 TRUE / error flag, TRUE on fault-level eErr
    bValid           : BOOL;                  // 返回值是否可用（故障级为 FALSE）/ return usable, FALSE on fault level
END_VAR
VAR CONSTANT
    DL_DATE_DAYS_MIN : DINT := 0;             // 纪元日，天数下界 [日] / the epoch day, lower bound [day]
    DL_DATE_DAYS_MAX : DINT := 65535;         // 保守容器口径上限，无符号 16 位天数顶 [日] / conservative container top, unsigned 16-bit day limit [day]
    DL_EPOCH_DATE_ZERO : DATE := DATE#1970-01-01; // 纪元起始日期 / the epoch date
    DL_DINT_ZERO     : DINT := 0;             // 有符号零常量，避免裸字面量 [日] / signed zero constant [day]
END_VAR
VAR
    nDays            : DINT;                  // 自纪元起天数中间量 [日] / day count intermediate since the epoch [day]
END_VAR

// 段 1｜返回值与错误状态预置 / segment 1, preset return value and error status
FC_DL_DateToDintDays := DL_DINT_ZERO;         // 故障缺省返回 0 [日] / fault default returns zero [day]
eErr := 0;                                    // 预置无错误 / preset no error
bError := FALSE;                              // 预置无故障 / preset no fault
bValid := FALSE;                              // 预置不可用，通过闸门后置位 / preset invalid, set TRUE after the gates
nDays := DL_DINT_ZERO;                        // 中间量清零 / clear the intermediate

// 段 2｜下域闸门：早于纪元的日期先于内建拦下 / segment 2, epoch lower gate precedes the built-in call
IF dateIn < DL_EPOCH_DATE_ZERO THEN
    eErr := 16#0001_0336;                     // 故障级：输入早于纪元 / fault level, the input precedes the epoch
    bError := TRUE;                           // 置故障标志 / raise the error flag
    bValid := FALSE;                          // 返回值不可用 / flag the return as unusable
    FC_DL_DateToDintDays := DL_DINT_ZERO;     // 确定缺省值 0 / deterministic default of zero
    RETURN;                                   // 出口，不触碰内建 / exit, the built-in is never touched
END_IF

// 段 3｜主体：域内才委托平台内建（天数口径）/ segment 3, delegate the built-in only inside the domain
nDays := DATE_TO_DINT(dateIn);                // 内建换算：DATE → 自纪元天数 [日] / built-in conversion from DATE to days since the epoch [day]

// 段 4｜容器溢出闸：内建给负天数即平台 DATE 位型承载异常 / segment 4, container overflow gate
IF nDays < DL_DATE_DAYS_MIN THEN
    eErr := 16#0001_0337;                     // 故障级：DATE 非法或容器溢出 / fault level, illegal DATE or container overflow
    bError := TRUE;                           // 置故障标志 / raise the error flag
    bValid := FALSE;                          // 返回值不可用 / flag the return as unusable
    FC_DL_DateToDintDays := DL_DINT_ZERO;     // 确定缺省值 0 / deterministic default of zero
    RETURN;                                   // 出口 / exit
END_IF

// 段 5｜保守容器口径钳位（信息级，钳位事件必须可见）/ segment 5, conservative container clamp at info level
IF nDays > DL_DATE_DAYS_MAX THEN
    nDays := DL_DATE_DAYS_MAX;                // 钳位至容器顶 [日] / clamp to the container top [day]
    eErr := 16#0001_0410;                     // 信息级：超保守口径已钳位，值仍可用 / info level, clamped to the conservative top, still usable
END_IF

// 段 6｜发布结果 / segment 6, publish the result
FC_DL_DateToDintDays := nDays;                // 输出自纪元起天数 [日] / publish the days since the epoch [day]
bValid := TRUE;                               // 域内或已钳位均可用 / usable in domain or after the clamp
END_FUNCTION

(* ---- FC_DL_DateToIsoString.st ---- *)
(*
    组件名称 : FC_DL_DateToIsoString
    所属子库 : DL_MathData
    当前版本 : 1.0.1
    兼 容 性 : CODESYS V3.5+ / TwinCAT 3 / 汇川 InoProShop；仅依赖 Standard.library
    功能描述 : DATE → 'YYYY-MM-DD' 十字符定宽文本，同时把年/月/日分解结果单出口，供 MES 台账与文件名直接取用。
              取舍 ①：用 Howard Hinnant 的 civil_from_days 整数算法反算日历 —— 纯整数、无查表、无浮点、无循环，
              对任意天数一次算到位；相比「按年循环扣天数」的写法，没有循环也就没有死循环风险与扫描周期抖动。
              取舍 ②：回代自校验（days_from_civil 反算天数必须等于输入）—— 日期算法的错误往往表现为「差一天」，
              这种错在报表上极难发现，回代一次就能把「算法实现错」与「输入数据错」彻底分开；
              自校验不过就绝不输出日期。
              取舍 ③：不做平台 DATE_TO_DTL 委托 —— DTL 结构体在部分平台的字段宽度与日期语义不一致，
              且本件只需要三个整数；直接走 DATE_TO_DINT 天数口径，链路最短。
              取舍 ④：早于纪元（1970-01-01）一律判故障 —— 负数天数在部分平台 DATE 实现里是「不支持」而非「负日期」，
              与其猜，不如让调用方知道这个值不可信。
    开源溯源 : T2-1 LGF Converter 子族（只借「日期转定宽文本」这一行为定义）。civil_from_days / days_from_civil；本件为道莅 clean-room 防御性实现（仅借 LGF 分类事实/参数域/行为定义，零代码行与符号名复制）。
              为公开算法（Howard Hinnant，公有领域），本实现按整数语义重写，零代码行与注释复制；
              码位、错误分级、自校验策略 100% 自有。
    本文件内含 : FUNCTION FC_DL_DateToIsoString（单 POU，无配套类型）
    依 赖 : 无 DL_ 内部依赖；Standard.library: LEN / MID / CONCAT
    红线自检 : R1 ✓ 零全局变量与外部变量 ｜ R2 ✓ 零物理 IO 地址
              R3 ✓ 纯 IEC 61131-3 ｜ R4 ✓ 纪元闸 + 年份域闸 + 回代自校验 + 输出长度自证（全整数，无除法零风险）
              R5 ✓ 全变量中英双语同行注释 ｜ R6 N/A 纯函数无顺序状态机，无 CASE 可写
              R7 N/A 无定时器、无沿检测实例 ｜ R8 ✓ 纪元常数、闰年基数、月长基数全常量化
    错误码   : 16#0001_0450 [信息级] 输出串长异常（补零逻辑防御提示），bValid = TRUE
               16#0001_0451 [信息级] 预留禁用（不得挪用）
               16#0001_0396 [故障级] 早于纪元或年份越 1970~9999，返回 '1970-01-01'，bValid = FALSE
               16#0001_0397 [故障级] 回代自校验失败（算法自证不过），返回 '1970-01-01'，bValid = FALSE
               16#0001_0398 [故障级] 预留禁用（不得挪用）
    码位总账 : 16#0001_0450 用 / 16#0001_0451 预留 ｜ 16#0001_0396 用 / 16#0001_0397 用 / 16#0001_0398 预留
    遗留假设 : ① 【编译门槛未闭合】本件依赖「DATE_TO_DINT 返回自 1970-01-01 起的天数、纪元当日记 0」这一口径。
              CODESYS / TwinCAT 3 默认如此，InoProShop 未实测；若某平台返回秒或返回 1970-01-01 记 1，
              回代自校验会失败并置 0397（可观测，不会静默出错）。
              ② 整数除法在三平台均向零截断，本件全部操作数为非负，故截断方向不敏感 —— IEC 语义推导，未逐平台实测。
              ③ MID 参数序按 IEC 标准 MID(串, 长度, 位置)，与库内既有用法同序。
    修订历史 :
        2026-11-16  v1.0.0  首版，R21 批次 3 入库
        2026-11-16  v1.0.1  R21 终审修复（严重）：年序判据末项除数误用 DL_ERA_DAYS = 146097，
                            而 Hinnant civil_from_days 该处应为「周期内最大天序」146096。二者仅在
                            nDoe = 146096（即每个 400 年周期的最后一天 = 世纪闰日 2 月 29 日）时结果不同：
                            错值使 nYoe = 400 越出 [0, 399]，回代自校验随即失败，2000-02-29 / 2400-02-29
                            等合法日期被误判为 0397 故障并回退成 '1970-01-01'。新增常量 DL_ERA_LAST = 146096
                            并改用于该式；其余天序取值两种除数同解，故本次修复零副作用。向量已用等价脚本
                            复算：1970-01-01 / 1999-12-31 / 2000-02-29 / 2026-11-16 / 9999-12-31 全部自校验通过。
*)
FUNCTION FC_DL_DateToIsoString : STRING
VAR_INPUT
    dateIn          : DATE;   // 待格式化日期，有效域 1970-01-01 ~ 9999-12-31 / date to format, valid from 1970-01-01 to 9999-12-31
END_VAR
VAR_OUTPUT
    eErr            : UDINT;  // 错误码，0=正常；16#0001_04XX 信息级 / 16#0001_03XX 故障级 / error id, 0=ok
    bError          : BOOL;   // 故障级标志，eErr 落 16#0001_03XX 时为 TRUE / fault flag, TRUE on fault-level eErr
    bValid          : BOOL;   // 返回值是否可用 / result usable flag
    nYear           : INT;    // 分解出的年份 1970~9999 [年] / decomposed year [year]
    nMonth          : INT;    // 分解出的月份 1~12 [月] / decomposed month [month]
    nDay            : INT;    // 分解出的日 1~31 [日] / decomposed day [day]
END_VAR
VAR
    nDays           : DINT;   // 自纪元起的天数 [天] / days since the epoch [day]
    nZ              : DINT;   // 纪元平移后的天数（+719468）[天] / day count shifted by the epoch offset [day]
    nEra            : DINT;   // 400 年周期序号 [周期] / four hundred year era index [era]
    nDoe            : DINT;   // 纪元年内的天序 0~146096 [天] / day of era, 0..146096 [day]
    nYoe            : DINT;   // 纪元年内年序 0~399 [年] / year of era, 0..399 [year]
    nDoy            : DINT;   // 年内的天序 0~365 [天] / day of year, 0..365 [day]
    nMp             : DINT;   // 三月起算的月序 0~11 [月] / month index counted from March, 0..11 [month]
    nY              : DINT;   // 工作年值 [年] / working year value [year]
    nM              : DINT;   // 工作月值 [月] / working month value [month]
    nD              : DINT;   // 工作日值 [日] / working day value [day]
    nCheck          : DINT;   // 回代算出的天数，用于自校验 [天] / recomputed day count used for the self check [day]
    nChkY           : DINT;   // 回代用年 [年] / year used by the reverse pass [year]
    nChkYoe         : DINT;   // 回代纪元年内年序 0~399 [年] / year of era used by the reverse pass [year]
    nChkDoy         : DINT;   // 回代用年内天序 [天] / day of year used by the reverse pass [day]
    nChkDoe         : DINT;   // 回代用纪元年内天序 [天] / day of era used by the reverse pass [day]
    sRet            : STRING; // 结果装配缓冲 [字符] / result assembly buffer [char]
    nLen            : INT;    // 结果实际长度 [字符] / actual result length [char]
END_VAR
VAR CONSTANT
    DL_ISO_LEN          : INT := 10;                 // 目标串长 'YYYY-MM-DD' [字符] / target length [char]
    DL_EPOCH_YEAR       : INT := 1970;               // 纪元年份 [年] / epoch year [year]
    DL_YEAR_MIN         : INT := 1970;               // 年份下界 [年] / lower year bound [year]
    DL_YEAR_MAX         : INT := 9999;               // 年份上界 [年] / upper year bound [year]
    DL_EPOCH_OFFSET     : DINT := 719468;            // 1970-01-01 在 Hinnant 纪元中的天序 [天] / epoch offset of 1970-01-01 [day]
    DL_ERA_DAYS         : DINT := 146097;            // 400 年周期的天数 [天] / days in a four hundred year era [day]
    DL_ERA_LAST         : DINT := 146096;            // 400 年周期内最大天序 = DL_ERA_DAYS − 1，年序判据专用除数 [天] / last day index inside an era, the dedicated divisor of the year-of-era test [day]
    DL_ERA_YEARS        : DINT := 400;               // 400 年周期的年数 [年] / years in an era [year]
    DL_CENTURY_DAYS     : DINT := 36524;             // 百年天数（闰日扣除用）[天] / days in a century used by the leap correction [day]
    DL_QUAD_DAYS        : DINT := 1460;              // 四年天数（闰日扣除用）[天] / days in four years used by the leap correction [day]
    DL_CENTURY_YEARS    : DINT := 100;               // 百年年数 [年] / years in a century [year]
    DL_YEAR_DAYS        : DINT := 365;               // 平年天数 [天] / days in a common year [day]
    DL_LEAP_DIV         : DINT := 4;                 // 四年闰基数 [年] / four year leap radix [year]
    DL_MONTH_SHIFT      : DINT := 3;                 // 三月起算的月偏移 [月] / month shift of the March based calendar [month]
    DL_MONTH_BASE       : DINT := 10;                // 三月起算的月份分界 [月] / boundary between the two month groups [month]
    DL_MONTH_ROLL       : DINT := 9;                 // 月份回卷量（mp + 3 − 12）[月] / month roll over amount [month]
    DL_MONTH_SUB        : DINT := 3;                 // 回代时 m > 2 分支的月偏移量（m − 3）[月] / month offset of the m greater than two branch [month]
    DL_MONTH_FEB        : DINT := 2;                 // 一、二月的分界值 [月] / boundary value of January and February [month]
    DL_DOY_SCALE        : DINT := 153;               // 月长累加系数 153 = 5 个月 × 30.6 [无量纲] / month length coefficient [dimensionless]
    DL_DOY_BIAS         : DINT := 2;                 // 月序取整偏置 [无量纲] / rounding bias of the month index [dimensionless]
    DL_DOY_DIV          : DINT := 5;                 // 月序除数 [无量纲] / divisor of the month index [dimensionless]
    DL_DIGIT_TABLE      : STRING := '0123456789';    // 数字字符表，MID 位置 = 值 + 1 [字符] / digit table, the MID position is the value plus one [char]
    DL_ISO_DASH         : STRING := '-';             // 日期分隔符 [字符] / date separator [char]
    DL_ISO_FALLBACK     : STRING := '1970-01-01';    // 故障回退串，长度恒 10 [字符] / fault fallback text with a constant length of ten [char]
    DL_ISO_ONE          : INT := 1;                  // 单位哨兵，MID 位置 1 基 [无量纲] / unity sentinel, MID is one based [dimensionless]
    DL_ISO_DIGIT_TEN    : DINT := 10;                // 十进制位数基数 [无量纲] / decimal digit radix [dimensionless]
    DL_ISO_DIGIT_HUND   : DINT := 100;               // 百位基数 [无量纲] / hundreds radix [dimensionless]
    DL_ISO_DIGIT_THOU   : DINT := 1000;              // 千位基数 [无量纲] / thousands radix [dimensionless]
    DL_DINT_ZERO        : DINT := 0;                 // 零哨兵 [无量纲] / zero sentinel [dimensionless]
    DL_INT_ZERO         : INT := 0;                  // 整数零哨兵，月份判零用 [月] / integer zero sentinel [month]
    DL_ERR_NONE         : UDINT := 16#0000_0000;     // 无故障 / no error
END_VAR

// 段 1｜返回值与错误状态预置 / segment 1, preset the return value and the error state
FC_DL_DateToIsoString := DL_ISO_FALLBACK;   // 故障缺省返回纪元日 / fault default returns the epoch date
eErr   := DL_ERR_NONE;                       // 预置无错误 / preset no error
bError := FALSE;                             // 预置无故障 / preset no fault
bValid := FALSE;                             // 预置结果不可用 / preset unusable
nYear  := DL_EPOCH_YEAR;                     // 预置年份为纪元年 / preset the year to the epoch
nMonth := 1;                                 // 预置月 1 / preset the month to one
nDay   := 1;                                 // 预置日 1 / preset the day to one
sRet   := '';                                // 缓冲清空 / clear the buffer

// 段 2｜天数口径与纪元闸 / segment 2, day count and epoch gate
nDays := DATE_TO_DINT(dateIn);               // 天数口径（1970-01-01 = 0），见遗留假设 ① / day count with the epoch at zero, see assumption one
IF nDays < DL_DINT_ZERO THEN
    eErr   := 16#0001_0396;                  // 早于纪元（故障级）/ earlier than the epoch, fault level
    bError := TRUE;                          // 置故障标志 / raise the fault flag
    RETURN;                                  // 返回纪元日 / return the epoch date
END_IF

// 段 3｜civil_from_days 反算（全整数，无循环）/ segment 3, civil from days with integer arithmetic only
nZ    := nDays + DL_EPOCH_OFFSET;            // 平移到 Hinnant 纪元 / shift into the Hinnant epoch
nEra  := nZ / DL_ERA_DAYS;                   // nZ 恒为正，直接整除即可 / nZ is always positive, a plain division suffices
nDoe  := nZ - nEra * DL_ERA_DAYS;            // 纪元年内天序 / day of era
nYoe  := (nDoe - nDoe / DL_QUAD_DAYS + nDoe / DL_CENTURY_DAYS - nDoe / DL_ERA_LAST) / DL_YEAR_DAYS;   // 纪元年内年序，末项除数为 146096 而非 146097 / year of era, the last divisor is 146096 not 146097
nY    := nYoe + nEra * DL_ERA_YEARS;         // 绝对年份 / absolute year
nDoy  := nDoe - (DL_YEAR_DAYS * nYoe + nYoe / DL_LEAP_DIV - nYoe / DL_CENTURY_YEARS);                 // 年内天序 / day of year
nMp   := (DL_DOY_DIV * nDoy + DL_DOY_BIAS) / DL_DOY_SCALE;                                            // 三月起算月序 / March based month index
nD    := nDoy - (DL_DOY_SCALE * nMp + DL_DOY_BIAS) / DL_DOY_DIV + DL_ISO_ONE;                         // 日 / day of month
IF nMp < DL_MONTH_BASE THEN
    nM := nMp + DL_MONTH_SHIFT;              // 三月到十二月 / March to December
ELSE
    nM := nMp - DL_MONTH_ROLL;               // 一月与二月，顺带年前推已在下面补 / January and February
END_IF
IF nM <= DL_MONTH_FEB THEN
    nY := nY + DL_ISO_ONE;                   // 一、二月属上一日历年，年值补一 / January and February belong to the previous calendar year
END_IF

// 段 4｜年份域闸 / segment 4, year domain gate
IF (nY < DL_YEAR_MIN) OR (nY > DL_YEAR_MAX) THEN
    eErr   := 16#0001_0396;                  // 年份越域（故障级）/ year out of domain, fault level
    bError := TRUE;                          // 置故障标志 / raise the fault flag
    RETURN;                                  // 返回纪元日 / return the epoch date
END_IF

// 段 5｜回代自校验：days_from_civil(y, m, d) 必须等于输入天数 / segment 5, reverse self check
nChkY := nY;                                 // 回代用年，取分解结果 / reverse pass year taken from the decomposed result
IF nM <= DL_MONTH_FEB THEN
    nChkY := nChkY - DL_ISO_ONE;             // 一、二月回退一年 / January and February roll the year back
END_IF
IF nM > DL_MONTH_FEB THEN
    nChkDoy := (DL_DOY_SCALE * (nM - DL_MONTH_SUB) + DL_DOY_BIAS) / DL_DOY_DIV + nD - DL_ISO_ONE;   // 三月起算的天序 / day of year for the March based branch
ELSE
    nChkDoy := (DL_DOY_SCALE * (nM + DL_MONTH_ROLL) + DL_DOY_BIAS) / DL_DOY_DIV + nD - DL_ISO_ONE;   // 一、二月的天序 / day of year for January and February
END_IF
nChkYoe := nChkY - (nChkY / DL_ERA_YEARS) * DL_ERA_YEARS;                                              // 纪元年内年序 0~399 / year of era
nChkDoe := nChkYoe * DL_YEAR_DAYS + nChkYoe / DL_LEAP_DIV - nChkYoe / DL_CENTURY_YEARS + nChkDoy;      // 年内闰日修正后加天序 / leap corrected day of year
nCheck  := (nChkY / DL_ERA_YEARS) * DL_ERA_DAYS + nChkDoe - DL_EPOCH_OFFSET;                            // 回代天数 / recomputed day count
IF nCheck <> nDays THEN
    eErr   := 16#0001_0397;                  // 回代自校验失败（故障级）/ reverse self check failed, fault level
    bError := TRUE;                          // 置故障标志 / raise the fault flag
    RETURN;                                  // 不输出未经复验的日期 / never publish an unverified date
END_IF

// 段 6｜定宽格式化：年 4 位、月日 2 位，逐位查表 / segment 6, fixed width formatting with table lookups
sRet := CONCAT(sRet, MID(DL_DIGIT_TABLE, DL_ISO_ONE, DINT_TO_INT(nY / DL_ISO_DIGIT_THOU) + DL_ISO_ONE));                                  // 千位 / thousands
sRet := CONCAT(sRet, MID(DL_DIGIT_TABLE, DL_ISO_ONE, DINT_TO_INT((nY / DL_ISO_DIGIT_HUND) MOD DL_ISO_DIGIT_TEN) + DL_ISO_ONE));           // 百位 / hundreds
sRet := CONCAT(sRet, MID(DL_DIGIT_TABLE, DL_ISO_ONE, DINT_TO_INT((nY / DL_ISO_DIGIT_TEN) MOD DL_ISO_DIGIT_TEN) + DL_ISO_ONE));            // 十位 / tens
sRet := CONCAT(sRet, MID(DL_DIGIT_TABLE, DL_ISO_ONE, DINT_TO_INT(nY MOD DL_ISO_DIGIT_TEN) + DL_ISO_ONE));                                 // 个位 / units
sRet := CONCAT(sRet, DL_ISO_DASH);           // 分隔符 / separator
sRet := CONCAT(sRet, MID(DL_DIGIT_TABLE, DL_ISO_ONE, DINT_TO_INT(nM / DL_ISO_DIGIT_TEN) + DL_ISO_ONE));                                   // 月十位 / month tens
sRet := CONCAT(sRet, MID(DL_DIGIT_TABLE, DL_ISO_ONE, DINT_TO_INT(nM MOD DL_ISO_DIGIT_TEN) + DL_ISO_ONE));                                 // 月个位 / month units
sRet := CONCAT(sRet, DL_ISO_DASH);           // 分隔符 / separator
sRet := CONCAT(sRet, MID(DL_DIGIT_TABLE, DL_ISO_ONE, DINT_TO_INT(nD / DL_ISO_DIGIT_TEN) + DL_ISO_ONE));                                   // 日十位 / day tens
sRet := CONCAT(sRet, MID(DL_DIGIT_TABLE, DL_ISO_ONE, DINT_TO_INT(nD MOD DL_ISO_DIGIT_TEN) + DL_ISO_ONE));                                 // 日个位 / day units

// 段 7｜分解结果单出口与长度自证 / segment 7, decomposed values and length self proof
nYear  := DINT_TO_INT(nY);                   // 年份出口 / publish the year
nMonth := DINT_TO_INT(nM);                   // 月份出口 / publish the month
nDay   := DINT_TO_INT(nD);                   // 日出口 / publish the day
nLen   := LEN(sRet);                         // 实际长度 / the actual length
IF nLen <> DL_ISO_LEN THEN
    eErr := 16#0001_0450;                    // 输出串长异常（信息级，只提示补零逻辑异常）/ length anomaly, info level
END_IF

// 段 8｜出口 / segment 8, exit
FC_DL_DateToIsoString := sRet;               // 输出 ISO 日期文本 / publish the ISO date text
bValid := TRUE;                              // 结果可用 / the result is usable
END_FUNCTION

(* ---- FC_DL_Deadband.st ---- *)
(*==============================================================================
 * 组件名称 (Component)  : FC_DL_Deadband
 * 所属子库 (Sublibrary) : DL_MathData
 * 当前版本 (Version)    : 1.0.0
 * 兼容性   (Platform)   : CODESYS 3.5 / TwinCAT 3 / 汇川 InoProShop / Machine Expert
 *                         仅依赖 Standard.library（ABS），全 REAL 运算
 * 功能描述 (Function)   : 死区（Dead Band）处理，用于抑制零点附近的传感器零漂、
 *                         量化噪声与计算残差，典型用途是 PID 误差通道，防止调节阀
 *                         在设定点附近高频动作导致定位器磨损。
 *                         提供两种互斥语义（由 bZeroMode 选择，不可同时生效）：
 *                         移位型（默认）：死区内输出 0，死区外输出 dev - sign(dev)*width，
 *                                        边界连续、无阶跃，可串入闭环；
 *                         归零型：死区内输出 0，死区外原样输出 dev，
 *                                边界有跳变（跳变量 = 死区宽度），属阈值开关直觉。
 * 失真披露 (Distortion): 死区必然使信号失真，失真量恰为死区宽度。用于 PID 误差通道时
 *                         fCenter 必须为 0，否则零点被人工搬移，积分项会持续累积偏置。
 * 开源溯源 (Origin)     : 原创实现。限幅思想参考 OSCAT DEAD_BAND_A 的 LM 处理，
 *                         语义与故障码按本库体系重写，未复制源码。
 * 依赖     (Depends)    : 无 DL_ 内部依赖
 * 红线自检 (Redline)    : R1 ✓ 零全局变量表与外部变量引用 ｜ R2 ✓ 零物理 IO 地址直写
 *                         R3 ✓ 纯 IEC 61131-3（自建符号函数，无标准 SIGN）
 *                         R4 ✓ 负宽容错 / 零宽直通 / 浮点容差 / 宽度上限
 *                         R5 ✓ 全变量中英双语同行注释 ｜ R6 N/A（无状态机）｜ R7 N/A（无实例调用）
 * 修订历史 (Revision)   :
 *   2026-11-14  v1.0.0  首版入库（Phase 1 冷启动 · Level 0 批次）
 *============================================================================*)
FUNCTION FC_DL_Deadband : REAL
VAR_INPUT
    fIn       : REAL;              // 输入值 [EU] / Input value [EU]
    fWidth    : REAL := 0.0;       // 死区半宽 [EU]，负值取绝对值 / Deadband half-width [EU], negative taken as absolute
    fCenter   : REAL := 0.0;       // 死区中心偏移 [EU]，零点不在 0 时使用 / Deadband center offset [EU]
    bZeroMode : BOOL := FALSE;     // FALSE = 移位型（连续），TRUE = 归零型（阈值开关） / FALSE = shift type, TRUE = zero type
END_VAR
VAR_OUTPUT
    bInDeadband : BOOL;            // 当前处于死区内 / Currently inside the deadband
    fDeviation  : REAL;            // 去中心后的原始偏差 [EU] / Raw deviation from the center [EU]
    fEffWidth   : REAL;            // 实际生效的死区半宽 [EU] / Effective deadband half-width [EU]
    uErrorId    : UDINT;           // 故障码，0 = 无故障 / Error code, 0 = no error
END_VAR
VAR
    fSign       : REAL;            // 自建符号函数结果，取值 +1.0 或 -1.0 / Self-built sign result, +1.0 or -1.0
    fWidthAbs   : REAL;            // 原始宽度的绝对值 [EU] / Absolute value of the input width [EU]
END_VAR
VAR CONSTANT
    DL_FLOAT_EPS      : REAL := 1.0E-6;      // 浮点判零容差 / Float zero tolerance
    DL_DEADBAND_MAX_WIDTH : REAL := 1000.0;  // 死区半宽硬上限 [EU]，防参数误填成 999 导致输出恒 0 / Hard upper limit [EU]
END_VAR

(*------------------------------------------------------------------------------
 * 段 1｜安全预置：返回值先落到"直通"语义，异常路径不引入额外失真
 *      Safe preset: default to pass-through so error paths add no extra distortion
 *-----------------------------------------------------------------------------*)
FC_DL_Deadband := fIn;
bInDeadband    := FALSE;
fDeviation     := 0.0;
fEffWidth      := 0.0;
fSign          := 1.0;
fWidthAbs      := 0.0;
uErrorId       := 16#0000_0000;

(*------------------------------------------------------------------------------
 * 段 2｜负宽度容错（边界 B1）：取绝对值后继续运行，绝不把宽度压成 0
 *      Negative width tolerance: take the absolute value and keep running
 *      宽度为 0 等价于死区消失，阀门会立刻恢复高频动作，正是现场最怕的结果，
 *      因此这里只告警、不降级
 *-----------------------------------------------------------------------------*)
fWidthAbs := ABS(fWidth);
fEffWidth := fWidthAbs;

IF fWidth < 0.0 THEN
    uErrorId := 16#0001_0003;
END_IF

(*------------------------------------------------------------------------------
 * 段 3｜宽度上限保护（边界 B5）：防止参数误填导致输出恒为 0
 *      Width upper limit: prevents a mis-typed parameter from freezing the output at 0
 *      "输出恒 0"在现场表现为"设备不响应"而非"参数错误"，极难定位，
 *      因此宁可钳位并告警，也要保证回路仍有响应
 *-----------------------------------------------------------------------------*)
IF fEffWidth > DL_DEADBAND_MAX_WIDTH THEN
    fEffWidth := DL_DEADBAND_MAX_WIDTH;
    uErrorId  := 16#0001_0003;
END_IF

(*------------------------------------------------------------------------------
 * 段 4｜偏差计算：先去掉中心偏移，后续所有判定只基于 fDeviation
 *      Deviation computation: remove the center offset first, all tests use fDeviation
 *-----------------------------------------------------------------------------*)
fDeviation := fIn - fCenter;

(*------------------------------------------------------------------------------
 * 段 5｜零宽度直通（边界 B2/B4）：严格直通，且不判为"在死区内"
 *      Zero-width pass-through: strict pass-through, never reported as inside the band
 *      判定用 ABS(..) <= EPS 的容差比较，禁止 fEffWidth = 0.0
 *-----------------------------------------------------------------------------*)
IF fEffWidth <= DL_FLOAT_EPS THEN
    FC_DL_Deadband := fDeviation;
    bInDeadband    := FALSE;
    RETURN;
END_IF

(*------------------------------------------------------------------------------
 * 段 6｜死区内判定：使用严格小于，边界点算"死区外"，保证移位型在边界连续
 *      Inside-band test: strict less-than keeps the shift type continuous at the edge
 *-----------------------------------------------------------------------------*)
IF ABS(fDeviation) < fEffWidth THEN
    bInDeadband    := TRUE;
    FC_DL_Deadband := 0.0;
ELSE
    IF bZeroMode THEN
        (*----------------------------------------------------------------------
         * 段 7a｜归零型：死区外原样输出，边界处存在等于死区宽度的阶跃
         *       Zero type: pass the deviation through, step size equals the band width
         *---------------------------------------------------------------------*)
        FC_DL_Deadband := fDeviation;
    ELSE
        (*----------------------------------------------------------------------
         * 段 7b｜移位型（默认）：减去带符号的死区宽度，边界连续无阶跃
         *       Shift type (default): subtract the signed band width, edge is continuous
         *       IEC 61131-3 无标准 SIGN 函数，必须自建；偏差为 0 时符号取 +1.0
         *       （此时实际不可达，因为已在段 6 判为死区内，仍显式给定以避免
         *        0/0 式未定义推导）
         *---------------------------------------------------------------------*)
        IF fDeviation >= 0.0 THEN
            fSign := 1.0;
        ELSE
            fSign := -1.0;
        END_IF

        FC_DL_Deadband := fDeviation - fSign * fEffWidth;
    END_IF
END_IF
END_FUNCTION

(* ---- FC_DL_DeburrBrushSpeedCalc.st ---- *)
(*
  DL Factory R88 | FC_DL_DeburrBrushSpeedCalc
  功能：算去毛刺刷丝线速度 v=π·D·n/60000 + vf·sinθ（进给修正项），超 25 m/s 报警
  开源溯源：无（clean-room 自研，依据公开工艺公式 刷轮线速度与进给投影叠加式，许可证=MIT，借鉴点=公式结构）
  规则：R1-R16 全遵守；R88 简单件标量形（纯标量入参出参，无循环体、无方法、无属性、无数组）
*)
FUNCTION FC_DL_DeburrBrushSpeedCalc : REAL
VAR_INPUT
    fDiaMm : REAL := 150.0; // 刷轮外径 D [mm] / brush wheel diameter [mm]
    fRpm : REAL := 2000.0; // 刷轮转速 n [r/min] / brush speed [rpm]
    fFeedMmPerS : REAL := 50.0; // 工件进给速度 vf [mm/s] / workpiece feed speed [mm/s]
    fContactDeg : REAL := 30.0; // 接触角 θ（刷丝与进给方向夹角，度制 0~90） [°] / contact angle in degrees [-]
    fLimitMPerS : REAL := 25.0; // 线速度报警阈值（刷丝飞散风险） [m/s] / overspeed alarm limit [m/s]
END_VAR
VAR_OUTPUT
    fSpeedMPerS : REAL; // 合成刷丝线速度 v [m/s] / resulting brush speed [m/s]
    xOverLimit : BOOL; // TRUE=线速度超过阈值，需报警 [-] / TRUE when above the alarm limit [-]
END_VAR
VAR
    fRotMPerS : REAL; // 旋转分量 π·D·n/60000 [m/s] / rotational component [m/s]
    fFeedMPerS : REAL; // 进给投影分量 vf·sinθ [m/s] / feed projection component [m/s]
    fAngleRad : REAL; // 接触角弧度值 [rad] / contact angle in radians [rad]
END_VAR

// 段 1｜出口预置
FC_DL_DeburrBrushSpeedCalc := -1.0; // 哨兵返回 -1（无效） [-] / sentinel return -1, invalid [-]
fSpeedMPerS := 0.0; // 合成线速度预置零 [m/s] / speed preset zero [m/s]
xOverLimit := FALSE; // 超限位预置 FALSE（未判定前不报超限） [-] / over-speed flag preset false [-]
fRotMPerS := 0.0; // 旋转分量预置零 [m/s] / rotational component preset zero [m/s]
fFeedMPerS := 0.0; // 进给分量预置零 [m/s] / feed component preset zero [m/s]
fAngleRad := 0.0; // 弧度预置零 [rad] / radians preset zero [rad]

// 段 2｜非有限拦截 + 域闸
IF NOT (fDiaMm > -1.0E30 AND fDiaMm < 1.0E30) OR NOT (fRpm > -1.0E30 AND fRpm < 1.0E30) THEN
    RETURN; // 直径/转速任一非有限即拒算 [-] / any non finite input rejected [-]
END_IF
IF NOT (fFeedMmPerS > -1.0E30 AND fFeedMmPerS < 1.0E30) OR NOT (fContactDeg > -1.0E30 AND fContactDeg < 1.0E30) THEN
    RETURN; // 进给/接触角任一非有限即拒算 [-] / any non finite input rejected [-]
END_IF
IF NOT (fLimitMPerS > -1.0E30 AND fLimitMPerS < 1.0E30) THEN
    RETURN; // 阈值非有限则报警判据失效，故先拦 [m/s] / the alarm limit must be finite [m/s]
END_IF
IF fDiaMm < 1.0E-9 OR fRpm < 0.0 OR fFeedMmPerS < 0.0 THEN
    RETURN; // 直径正域闸 + 转速/进给非负闸 [mm, r/min, mm/s] / positive diameter, non negative speeds
END_IF
IF fContactDeg < 0.0 OR fContactDeg > 90.0 THEN
    RETURN; // 接触角闭区间域闸 [0,90]，超界则 sinθ 投影无物理意义 [°] / contact angle closed interval gate [deg]
END_IF
IF fLimitMPerS <= 0.0 THEN
    RETURN; // 阈值正域闸：非正阈值会使报警恒真 [m/s] / positive limit gate [m/s]
END_IF

// 段 3｜计算
fAngleRad := fContactDeg * 0.0174532925; // 度 × (π/180) = rad，换算常数 0.0174532925 [rad] / degrees to radians [rad]
fRotMPerS := 3.14159265 * fDiaMm * fRpm / 60000.0; // mm × r/min ÷ 60000 = m/s；60000 恒正 [m/s] / rotational component [m/s]
fFeedMPerS := fFeedMmPerS * 0.001 * SIN(fAngleRad); // (mm/s) × 0.001 m/mm × [-] = m/s，进给投影项 [m/s] / [m/s]
fSpeedMPerS := fRotMPerS + fFeedMPerS; // m/s + m/s = m/s，两项合成 [m/s] / [m/s] + [m/s] = [m/s]

// 段 4｜判定与饱和
IF NOT (fSpeedMPerS > -1.0E30 AND fSpeedMPerS < 1.0E30) THEN
    RETURN; // 结果非有限再拦一次 [-] / re-check the result for finiteness [-]
END_IF
xOverLimit := fSpeedMPerS > fLimitMPerS; // 严格大于阈值为超限，等于阈值仍判合格 [m/s] / strict compare [m/s]

// 段 5｜出口自检
IF fSpeedMPerS < fRotMPerS THEN
    RETURN; // 出口自检：合成值不得小于旋转分量（说明叠加链被破坏） [m/s] / synthetic value must not drop below [m/s]
END_IF
FC_DL_DeburrBrushSpeedCalc := fSpeedMPerS; // 返回合成刷丝线速度 [m/s] / return the brush speed [m/s]
END_FUNCTION

(* ---- FC_DL_DegToRadEx.st ---- *)
(*
    FC_DL_DegToRadEx —— 度到弧度转换原子（LREAL 域）
    ------------------------------------------------------------------
    分类      : DL_MathData / Angle
    前缀      : FC_DL_
    版本      : 1.0.0
    溯源      : IEC 61131-3 标准语义的道莅防御性实现
                （内部委托乘法运算语义与 π 常数，外围统一错误码/钳位/双语文档；
                  未复制任何闭源厂商源码，参考实现仅限 MIT/Apache 许可）
    平台      : 纯 IEC 61131-3，CODESYS / TwinCAT / InoProShop 通用
    作者      : 道莅代码库 · PLC编程专家（R40）
    ------------------------------------------------------------------
    功能说明  : 度到弧度转换：返回 fDeg × (π / 180)，换算常数取 LREAL 精度
                字面量（≥16 位有效数字，R51 口径：REAL 精度常数禁入换算路径）；
                输入非有限（NaN 或 ±Inf）判为故障级 16#0001_03D0，返回 0.0 且
                bValid=FALSE（非有限值参与换算在三平台行为不一致，一律拦截）；
                溢出预判采用比较式消灭溢出路径（R54 口径：比较表达式内禁止出现
                乘法运算符，先判域后计算）：|fDeg| > LREAL 最大有限值 ÷ (π/180)
                时判乘积将溢出，判为故障级 16#0001_03D1，返回 0.0（不输出 Inf）；
                预判式除法合法性留档：换算常数 π/180 ≈ 0.017453292519943295 恒正
                且非零，除法本身无除零面；
                域内换算后再做结果非有限复检兜底（理论不可达：域闸后的乘积恒有限）。
    错误码    : 16#0001_03D0 输入非有限（NaN 或 ±Inf）——故障级，返回 0.0
                16#0001_03D1 换算乘积将溢出 LREAL 域（预判命中或复检失败）——故障级，返回 0.0
                （R90 反证句：溢出场景无法由输入非有限码观测——该场景输入有限而
                  结果非有限，与 16#0001_03D0 的「输入坏」语义无法区分，现有输出
                  组合无法还原「值大溢出」首因，故独立占码）
    非有限口径 : NaN 用自不等 f <> f，±Inf 用 (f − f) <> (f − f) 差值自减判定（R15）。
    状态机    : R6 标注 N/A —— 本组件为纯函数无顺序状态机，无 CASE 可写，
                非法状态不可能出现，故以本节说明替代 ELSE 兜底
    修订记录  : 2026-11-19 v1.0.0 首次入库（R40 · 批 2 · T0 快车道）
*)
FUNCTION FC_DL_DegToRadEx : LREAL
VAR_INPUT
    fDeg : LREAL; // 角度输入 [°] ｜ angle input in degrees
END_VAR
VAR_OUTPUT
    eErr   : UDINT; // 错误码，0=正常，16#0001_03XX=故障级 ｜ error id, 0=ok, 16#0001_03XX=fault level
    bError : BOOL;  // 是否出错，eErr 落故障级时为 TRUE ｜ fault flag, TRUE when eErr is fault level
    bValid : BOOL;  // 输出是否有效可用 ｜ output valid flag
END_VAR
VAR CONSTANT
    DL_DEG2RAD  : LREAL := 0.017453292519943295;      // 换算常数 π/180，LREAL 精度 ≥16 位有效数字 [rad/°] ｜ conversion constant pi/180, LREAL precision of at least 16 significant digits
    DL_LREAL_MAX: LREAL := 1.7976931348623157E308;    // LREAL 最大有限值 [无量纲] ｜ largest finite LREAL
END_VAR
VAR
    bNonFinite : BOOL; // 输入非有限判定结果 ｜ non-finite detection result of the input
    fOut       : LREAL; // 换算结果暂存，供出口复检 ｜ staging of the converted result for exit recheck
END_VAR

// 段 1｜返回值与错误状态预置 ｜ segment 1, preset return value and error status
FC_DL_DegToRadEx := 0.0; // 故障缺省返回 0 [rad] ｜ fault default returns 0
eErr   := 0;     // 预置无错误 ｜ preset no error
bError := FALSE; // 预置无故障 ｜ preset no fault
bValid := FALSE; // 预置无效，通过防御闸后置位 ｜ preset invalid, set TRUE after guard passes
fOut   := 0.0;   // 暂存清零 ｜ clear the staging value

// 段 2｜输入非有限防御闸（早退） ｜ segment 2, input non-finite guard (early return)
bNonFinite := (fDeg <> fDeg) OR ((fDeg - fDeg) <> (fDeg - fDeg)); // NaN 自不等 + 差值自减判 ±Inf [°] ｜ NaN by self-inequality, +/-Inf by self-subtraction
IF bNonFinite THEN
    FC_DL_DegToRadEx := 0.0; // 故障级返回 0 [rad] ｜ fault level returns 0
    eErr   := 16#0001_03D0;  // 输入非有限故障码 ｜ non-finite input fault id
    bError := TRUE;          // 置故障标志（R45 配对）｜ raise the fault flag (R45 pairing)
    bValid := FALSE;         // 输出无效 ｜ output invalid
    RETURN;                  // 早退 ｜ early return
END_IF

// 段 3｜溢出预判域闸（比较式，比较表达式内无乘法运算符） ｜ segment 3, overflow pre-check gate (comparison form, no multiplication inside the comparison)
IF ABS(fDeg) > (DL_LREAL_MAX / DL_DEG2RAD) THEN
    FC_DL_DegToRadEx := 0.0; // 预判命中不计算，返回 0 [rad] ｜ pre-check hit, no computation, returns 0
    eErr   := 16#0001_03D1;  // 换算溢出故障码 ｜ conversion overflow fault id
    bError := TRUE;          // 置故障标志（R45 配对）｜ raise the fault flag (R45 pairing)
    bValid := FALSE;         // 输出无效 ｜ output invalid
    RETURN;                  // 早退 ｜ early return
END_IF

// 段 4｜域内换算主体（末段） ｜ segment 4, in-domain conversion body (final)
fOut := fDeg * DL_DEG2RAD; // 度乘以换算常数得弧度 [rad] ｜ degrees times the conversion constant gives radians

// 段 5｜结果非有限复检兜底（理论不可达：域闸后的乘积恒有限） ｜ segment 5, result non-finite recheck (unreachable: the product after the gate is always finite)
IF (fOut <> fOut) OR ((fOut - fOut) <> (fOut - fOut)) THEN
    FC_DL_DegToRadEx := 0.0; // 复检失败按溢出处置 [rad] ｜ recheck failure treated as overflow
    eErr   := 16#0001_03D1;  // 复用溢出码（同因同码，不新占码位）｜ reuse the overflow code (same cause, no new code)
    bError := TRUE;          // 置故障标志 ｜ raise the fault flag
    bValid := FALSE;         // 输出无效 ｜ output invalid
    RETURN;                  // 早退 ｜ early return
END_IF

// 段 6｜出口装配 ｜ segment 6, exit assembly
FC_DL_DegToRadEx := fOut; // 换算结果直通 ｜ converted result pass-through
bError := FALSE;          // 正常出口不置故障 ｜ normal exit raises no fault
bValid := TRUE;           // 输出有效可用 ｜ output valid
END_FUNCTION

(* ---- FC_DL_DewPointSpreadCalc.st ---- *)
// FC_DL_DewPointSpreadCalc v1.0.0
(*==============================================================================
 * 功能描述: 露点温差计算。fSpreadK = 干球温度 - 露点温度 [K]；负值物理无效
 *           （露点不可能高于干球）→ bValid=FALSE 并返回饱和零域；任一输入非有限
 *           同样无效。
 * 接口契约: 输入 fTempC/fDewPointC [°C]；输出 bValid 回执，返回温差 [K]。
 * 修订历史: 2026-11-23  v1.0.0  R74 首版
 *==============================================================================*)

FUNCTION FC_DL_DewPointSpreadCalc : REAL
VAR_INPUT
    fTempC      : REAL := 20.0;   // 干球温度 [°C] / Dry-bulb temperature [degC]
    fDewPointC  : REAL := 10.0;   // 露点温度 [°C] / Dew-point temperature [degC]
END_VAR
VAR_OUTPUT
    bValid : BOOL;                // 结果有效回执 [-] / Result validity receipt
END_VAR

(* —— 段 0：全路径赋值缺省（无效安全侧） —— *)
bValid := FALSE;                             // 有效回执预清 / Validity preset
FC_DL_DewPointSpreadCalc := 0.0;             // 返回值缺省零 / Result default zero

(* —— 段 1：非有限闸（NaN 自反判） —— *)
IF (fTempC <> fTempC) OR (fDewPointC <> fDewPointC) THEN   // NaN 自反判（判等禁令唯一例外） / NaN self-reflexive tests
    RETURN;                                  // 无效返回零 / Invalid, return zero
END_IF

(* —— 段 2：温差换算与物理域校验（负温差判无效，浮点容差口径） —— *)
IF (fTempC - fDewPointC) < 0.0 THEN          // 负温差物理无效（露点高于干球） / Negative spread physically invalid
    RETURN;                                  // 无效返回零 / Invalid, return zero
END_IF
FC_DL_DewPointSpreadCalc := fTempC - fDewPointC;   // 露点温差 [K] / Dew-point spread [K]
bValid := TRUE;                              // 有效回执 / Validity receipt

END_FUNCTION

(* ---- FC_DL_DewPointToPpmV.st ---- *)
(*
  组件名 Component   : FC_DL_DewPointToPpmV
  子库 Sublibrary    : DL_MathData
  版本 Version       : 1.0.1
  兼容性 Platform    : CODESYS 3.5 / TwinCAT 3 / 汇川 InoProShop / Machine Expert（仅 Standard.library）
  功能 Function      : 露点温度 → 气体水分含量 ppmV 换算（饱和压比值法）：
                       1) 复用饱和蒸气压唯一属主 FC_DL_VaporPressureSat（DL_Algo）求露点温度
                       对应饱和水蒸气压 p_sat，本件零 Magnus 常数复制、零重复声明；
                       2) 摩尔分数 x_w = p_sat / p_total（分母总压前置正域判据，不进入除法）；
                       3) ppmV = x_w × 1E6，比值 > 1 时饱和钳位到 1.0 并置信息标志；
                       4) 非有限输入（NaN 自反判 + 无穷差值自减判）直接判无效返回 0.0。
  边界 Boundary      : ① 纯函数、无状态机、无内部实例，可重入；
                       ② 总压域 [1.0E-3, 2.0E7] Pa，域外判无效不外推；
                       ③ 露点温度域检查由属主承担，钳位标志透传（bClamped）；
                       ④ 无全局变量引用、无外部变量声明、无物理地址寻址；
                       ⑤ 结果仅当 bValid = TRUE 才可被工艺判据引用。
  依赖 Depends       : FC_DL_VaporPressureSat（DL_Algo，饱和压唯一属主，按 registry 实名调用）
  溯源 Origin        : 道莅自研 clean-room（参考 t2-1-lgf-converter 行为定义分类与参数域，
                       零代码行复制；饱和压计算完全委托既有属主）
  码位 Code          : 16#05_0_06
  码表 Error codes   : 纯函数件无状态机码轨；无效结果经 bValid = FALSE 表达（哨兵返回 0.0），
                       本件不占用故障码位（MathData 段 0005 内 0506 为本格独占声明，保留不用）。
  修订历史 Revision  :
    2026-11-19  v1.0.0  R44 首版（批次 1 · 序号 1）
    2026-11-23  v1.0.1  R73 补 bValid 回执：段 3 属主调用补收 bValid 局部回执，
                       回执无效并入既有哨兵零出口，契约不变
*)

FUNCTION FC_DL_DewPointToPpmV : LREAL
VAR_INPUT
    fDewPointC : LREAL;                 // 露点温度 [摄氏度]，域 -40.0..100.0（域检查属主承担）/ Dew point temperature
    fPressPa   : LREAL;                 // 气体总压 [Pa]，域 1.0E-3..2.0E7 / Total gas pressure
END_VAR
VAR_OUTPUT
    bValid     : BOOL;                  // 结果有效标志，FALSE 时返回值为哨兵 0.0 / Result validity flag
    bClamped   : BOOL;                  // 饱和压属主输入钳位标志透传 / Saturation owner clamped flag
    bSatRatio  : BOOL;                  // 比值超 1 已饱和钳位标志 / Ratio saturated and clamped flag
END_VAR
VAR
    fPsatPa   : LREAL;                  // 属主返回的饱和水蒸气压 [Pa] / Saturation vapor pressure from owner
    bSatOk    : BOOL;                   // 属主调用受理标志 / Owner call acceptance flag
    _bPwsValid: BOOL;                   // 属主输出可用回执 / Owner outputs-usable receipt
    _bPwsClamped : BOOL;    // 属主件钳位回执（本件不消费，仅契约全回执） / Owner clamp receipt (unused, full-receipt contract)
    _nPwsErr     : UDINT;   // 属主件错误码回执 / Owner error-code receipt
    _bPwsError   : BOOL;    // 属主件故障级回执 / Owner fault-flag receipt
END_VAR
VAR CONSTANT
    DL_PPM_SCALE : LREAL := 1.0E6;      // 摩尔分数 → ppmV 放大系数 [ppmV] / Mole fraction to ppmV scale
    DL_P_MIN     : LREAL := 1.0E-3;     // 总压有效下限 [Pa] / Pressure valid floor
    DL_P_MAX     : LREAL := 2.0E7;      // 总压有效上限 [Pa] / Pressure valid ceiling
    DL_RATIO_MAX : LREAL := 1.0;        // 摩尔分数物理上界 [无量纲] / Mole fraction physical ceiling
    DL_ZERO      : LREAL := 0.0;        // 无效哨兵返回值 [ppmV] / Sentinel return for invalid
END_VAR

(* —— 段 1｜出口预清零（纯函数无实例，无定时器/沿刷新义务） —— *)
bValid    := FALSE;                     // 缺省无效
bClamped  := FALSE;                     // 属主钳位标志缺省 FALSE
bSatRatio := FALSE;                     // 饱和钳位标志缺省 FALSE

(* —— 段 2｜输入防御：非有限值（NaN 自反 + 无穷差值自减）与总压域闸 —— *)
IF (fDewPointC <> fDewPointC) OR ((fDewPointC - fDewPointC) <> DL_ZERO)
   OR (fPressPa <> fPressPa) OR ((fPressPa - fPressPa) <> DL_ZERO)
   OR (fPressPa < DL_P_MIN) OR (fPressPa > DL_P_MAX) THEN
    FC_DL_DewPointToPpmV := DL_ZERO;    // 无效输入：哨兵零返回，不进入除法
    RETURN;
END_IF

(* —— 段 3｜委托饱和压唯一属主：禁在本件重复声明 Magnus 常数 —— *)
bSatOk := FC_DL_VaporPressureSat(fTempC := fDewPointC, fPvSat => fPsatPa, bClamped => bClamped, bValid => _bPwsValid, eErr => _nPwsErr, bError => _bPwsError);
IF (NOT bSatOk) OR (NOT _bPwsValid) THEN
    FC_DL_DewPointToPpmV := DL_ZERO;    // 属主判无效：哨兵零返回
    RETURN;
END_IF

(* —— 段 4｜饱和压比值法：分母已过正域闸，除法安全；比值超 1 饱和钳位 —— *)
IF fPsatPa > (fPressPa * DL_RATIO_MAX) THEN
    bSatRatio := TRUE;                  // 比值超物理上界：钳位并留痕
    FC_DL_DewPointToPpmV := DL_PPM_SCALE * DL_RATIO_MAX;
ELSE
    FC_DL_DewPointToPpmV := DL_PPM_SCALE * (fPsatPa / fPressPa);
END_IF
bValid := TRUE;                         // 全部防御通过：结果有效
END_FUNCTION

(* ---- FC_DL_DintDaysToDate.st ---- *)
(*
    FC_DL_DintDaysToDate —— 天数到 DATE 的还原
    ------------------------------------------------------------------
    分类      : DL_MathData / Convert
    前缀      : FC_DL_
    版本      : 1.0.0
    溯源      : IEC 61131-3 标准语义的道莅防御性实现（自 1970-01-01 起天数 → DATE）；
                委托平台内建 DINT_TO_DATE 完成还原，本件不重实现历法内核；
                域闸门、非饱和还原口径、错误分级与码位 100% 自有；
                clean-room 重写，未复制任何闭源厂商源码，参考实现仅限 MIT/Apache 许可
    平台      : 纯 IEC 61131-3，CODESYS V3.5+ / TwinCAT 3 / InoProShop 通用
    作者      : 道莅代码库 · PLC编程专家（R20）
    ------------------------------------------------------------------
    功能说明  : 把天数整型还原成日历日期，与 FC_DL_DateToDintDays 构成双向对。
                交付期、下次保养日、保质期到期日这类「数据库存天数、PLC 要日期」的场景，
                跨零点批量换算是高频口径。
                核心防御：① 负天数与超容器天数均返回纪元日并置 bValid = FALSE，
                   绝不做饱和还原——饱和会把越界天数改写成 1970-01-01 或容器顶，
                   台账上看不出异常，这是本件刻意与饱和族件分道的地方；
                ② 域端点（纪元日 0 与容器顶 65535）发信息级提示，便于排查上游哨兵值；
                ③ 天数上界与 FC_DL_DateToDintDays 用同一常量口径，正反两向不会错位。
                职责边界：日期天数化归 FC_DL_DateToDintDays；带偏移日期推算归
                FC_DL_DateAddDays（它先经天数路径再加偏移，天然覆盖本件域内域）。
    编译门槛  : 主路径依赖平台内建 DINT_TO_DATE（天数口径），三平台标准库均提供。
                若目标平台缺该内建，按「天数 → 纪元日零点 DT → DT 取日期」路径落地，
                中间量与闸门顺序不变；DL_DATE_DAYS_MAX 取 65535 保守口径，
                编码前按目标平台实测锚定（与 FC_DL_DateToDintDays 同源裁定）。
    错误码    : 16#0001_0412 天数恰为域端点（0 或 65535），已如实还原——信息级，值仍可用
                16#0001_0413 预留禁用（信息级，不得挪用）
                16#0001_0339 负天数（nDays < 0）——故障级，返回纪元日
                16#0001_033A 天数超容器域（nDays > 65535）——故障级，返回纪元日，不做饱和
                16#0001_033B 预留禁用（故障级，不得挪用）
    码位总账  : 16#0001_0412 用 / 16#0001_0413 预留 ｜ 16#0001_0339 用 / 16#0001_033A 用 / 16#0001_033B 预留
    状态机    : R6 标注 N/A —— 本组件为纯函数无顺序状态机，无 CASE 可写，非法状态不可能出现
    采样约定  : 本件无定时器、无沿检测、无状态；单拍纯计算，结论与任务周期无关。
    修订记录  : 2026-11-16 v1.0.0 首次入库（R20）
*)
FUNCTION FC_DL_DintDaysToDate : DATE
VAR_INPUT
    nDays            : DINT;                  // 自纪元起天数 [日]，有效域 0~65535 / days since the epoch [day], valid domain 0 to 65535
END_VAR
VAR_OUTPUT
    eErr             : UDINT;                 // 错误码，0=正常 / error id, 0=ok
    bError           : BOOL;                  // 故障标志，eErr 为故障级时 TRUE / error flag, TRUE on fault-level eErr
    bValid           : BOOL;                  // 返回值是否可用（故障级为 FALSE）/ return usable, FALSE on fault level
END_VAR
VAR CONSTANT
    DL_DATE_DAYS_MIN : DINT := 0;             // 纪元日，天数下界 [日] / the epoch day, lower bound [day]
    DL_DATE_DAYS_MAX : DINT := 65535;         // 保守容器口径上限，无符号 16 位天数顶 [日] / conservative container top, unsigned 16-bit day limit [day]
    DL_EPOCH_DATE_ZERO : DATE := DATE#1970-01-01; // 纪元起始日期，故障缺省返回 / the epoch date returned on faults
END_VAR
VAR
    nWork            : DINT;                  // 入参副本，避免改动调用方数据 [日] / input copy, never modifies caller data [day]
END_VAR

// 段 1｜返回值与错误状态预置 / segment 1, preset return value and error status
FC_DL_DintDaysToDate := DL_EPOCH_DATE_ZERO;   // 故障缺省返回纪元日 / fault default returns the epoch date
eErr := 0;                                    // 预置无错误 / preset no error
bError := FALSE;                              // 预置无故障 / preset no fault
bValid := FALSE;                              // 预置不可用，通过闸门后置位 / preset invalid, set TRUE after the gates
nWork := nDays;                               // 取入参副本参与判定 / copy the input for the comparisons

// 段 2｜下域闸门：负天数不是日期 / segment 2, negative gate, a negative day count is no date
IF nWork < DL_DATE_DAYS_MIN THEN
    eErr := 16#0001_0339;                     // 故障级：负天数 / fault level, negative day count
    bError := TRUE;                           // 置故障标志 / raise the error flag
    bValid := FALSE;                          // 返回值不可用 / flag the return as unusable
    RETURN;                                   // 出口，保持纪元日 / exit, the epoch date is kept
END_IF

// 段 3｜上域闸门：超容器域不做饱和（饱和会伪造日期）/ segment 3, upper gate without saturation
IF nWork > DL_DATE_DAYS_MAX THEN
    eErr := 16#0001_033A;                     // 故障级：超平台容器域 / fault level, beyond the platform container
    bError := TRUE;                           // 置故障标志 / raise the error flag
    bValid := FALSE;                          // 返回值不可用 / flag the return as unusable
    RETURN;                                   // 出口，保持纪元日，不伪造日期 / exit, no fabricated date
END_IF

// 段 4｜主体：域内才委托平台内建 / segment 4, delegate the built-in only inside the domain
FC_DL_DintDaysToDate := DINT_TO_DATE(nWork);  // 内建还原：天数 → 日期 / built-in conversion from days to a date
bValid := TRUE;                               // 域内还原可用 / the in-domain date is usable

// 段 5｜域端点提示（信息级，不置 bError）/ segment 5, domain endpoint hint at info level
IF (nWork = DL_DATE_DAYS_MIN) OR (nWork = DL_DATE_DAYS_MAX) THEN
    eErr := 16#0001_0412;                     // 信息级：天数恰为域端点，多为上游哨兵值 / info level, a domain endpoint, often an upstream sentinel
END_IF
END_FUNCTION

(* ---- FC_DL_DintEpochToDt.st ---- *)
(*
    FC_DL_DintEpochToDt —— Unix 纪元秒到 DATE_AND_TIME
    ------------------------------------------------------------------
    分类      : DL_MathData / Convert
    前缀      : FC_DL_
    版本      : 1.0.0
    溯源      : IEC 61131-3 标准语义的道莅防御性实现（Unix 纪元秒 → DATE_AND_TIME）；
                委托平台内建 DINT_TO_DT 完成还原，本件不重实现历法内核；
                域闸门、非饱和还原口径、错误分级与码位 100% 自有；
                clean-room 重写，未复制任何闭源厂商源码，参考实现仅限 MIT/Apache 许可
    平台      : 纯 IEC 61131-3，CODESYS V3.5+ / TwinCAT 3 / InoProShop 通用
    作者      : 道莅代码库 · PLC编程专家（R20）
    ------------------------------------------------------------------
    功能说明  : 把 MES / 日志侧回传的 Unix 纪元秒还原成 PLC 本地时刻，与
                FC_DL_DtToDintEpoch 构成双向对。
                核心防御：① 还原方向遇域外输入一律不输出「错值」——负秒与超 Y2038 秒
                   均返回纪元零点并置 bValid = FALSE，宁可不给时刻也不给错时刻，
                   因为错时刻会污染趋势曲线与批次记录，而空值只会触发一次重试；
                ② 本件不做饱和还原（与正向件的饱和出口刻意不同）：饱和会把数据库里的
                   越界秒静默改写成 2038-01-19，故障现场证据随之消失；
                ③ 边界秒（0 与 2147483647）发信息级提示，提示该值处于域端点，
                   便于排查上游把哨兵值当时刻下发的组态错。
                职责边界：正方向（DT → 纪元秒）归 FC_DL_DtToDintEpoch；
                本件只管「秒 → 时刻」单向还原。
    编译门槛  : 主路径依赖平台内建 DINT_TO_DT，三平台标准库均提供。
                若目标平台缺该内建，按合成路径落地：nDays = n / DL_SEC_PER_DAY、
                nSecOfDay = n MOD DL_SEC_PER_DAY，两操作数先判非负（段 2 已保证 n >= 0，
                余数口径安全），再 DINT_TO_DATE + DINT_TO_TOD 合成 DATE_AND_TIME。
                合成路径只在操作数非负域内使用模运算，与 TOD 回绕件的禁模纪律不冲突。
    错误码    : 16#0001_040E 输入恰为域端点（0 或 2147483647），已如实还原——信息级，值仍可用
                16#0001_040F 预留禁用（信息级，不得挪用）
                16#0001_0333 负纪元秒（nEpochSec < 0）——故障级，返回纪元零点
                16#0001_0334 超出 Y2038 秒域（nEpochSec > 2147483647）——故障级，返回纪元零点，不做饱和
                16#0001_0335 预留禁用（故障级，不得挪用）
    码位总账  : 16#0001_040E 用 / 16#0001_040F 预留 ｜ 16#0001_0333 用 / 16#0001_0334 用 / 16#0001_0335 预留
    状态机    : R6 标注 N/A —— 本组件为纯函数无顺序状态机，无 CASE 可写，非法状态不可能出现
    采样约定  : 本件无定时器、无沿检测、无状态；单拍纯计算，结论与任务周期无关。
    修订记录  : 2026-11-16 v1.0.0 首次入库（R20）
*)
FUNCTION FC_DL_DintEpochToDt : DATE_AND_TIME
VAR_INPUT
    nEpochSec        : DINT;                  // 纪元秒 [s]，有效域 0~2147483647 / epoch seconds [s], valid domain 0 to 2147483647
END_VAR
VAR_OUTPUT
    eErr             : UDINT;                 // 错误码，0=正常 / error id, 0=ok
    bError           : BOOL;                  // 故障标志，eErr 为故障级时 TRUE / error flag, TRUE on fault-level eErr
    bValid           : BOOL;                  // 返回值是否可用（故障级为 FALSE）/ return usable, FALSE on fault level
END_VAR
VAR CONSTANT
    DL_EPOCH_SEC_MAX : DINT := 2147483647;    // DINT 秒域上限，即 2038-01-19T03:14:07Z [s] / DINT second domain top, the Y2038 instant [s]
    DL_EPOCH_SEC_ZERO : DINT := 0;            // 纪元零点秒 [s] / the epoch second [s]
    DL_SEC_PER_DAY   : DINT := 86400;         // 每日秒数 [s/日]，合成路径的除数量 / seconds per day [s/day], divisor of the synthesis path
    DL_EPOCH_DT_ZERO : DATE_AND_TIME := DT#1970-01-01-00:00:00; // 纪元零点时刻，故障缺省返回 / the epoch instant returned on faults
END_VAR
VAR
    nWork            : DINT;                  // 入参副本，避免改动调用方数据 [s] / input copy, never modifies caller data [s]
END_VAR

// 段 1｜返回值与错误状态预置 / segment 1, preset return value and error status
FC_DL_DintEpochToDt := DL_EPOCH_DT_ZERO;      // 故障缺省返回纪元零点 / fault default returns the epoch instant
eErr := 0;                                    // 预置无错误 / preset no error
bError := FALSE;                              // 预置无故障 / preset no fault
bValid := FALSE;                              // 预置不可用，通过闸门后置位 / preset invalid, set TRUE after the gates
nWork := nEpochSec;                           // 取入参副本参与判定 / copy the input for the comparisons

// 段 2｜下域闸门：负秒不是时刻，绝不进内建 / segment 2, negative gate, a negative second is no instant
IF nWork < DL_EPOCH_SEC_ZERO THEN
    eErr := 16#0001_0333;                     // 故障级：负纪元秒 / fault level, negative epoch seconds
    bError := TRUE;                           // 置故障标志 / raise the error flag
    bValid := FALSE;                          // 返回值不可用 / flag the return as unusable
    RETURN;                                   // 出口，保持纪元零点 / exit, the epoch instant is kept
END_IF

// 段 3｜上域闸门：超 Y2038 域不做饱和（饱和会伪造时刻，破坏故障证据）/ segment 3, upper gate without saturation
IF nWork > DL_EPOCH_SEC_MAX THEN
    eErr := 16#0001_0334;                     // 故障级：超 Y2038 秒域 / fault level, beyond the Y2038 second domain
    bError := TRUE;                           // 置故障标志 / raise the error flag
    bValid := FALSE;                          // 返回值不可用 / flag the return as unusable
    RETURN;                                   // 出口，保持纪元零点，不伪造时刻 / exit, no fabricated instant
END_IF

// 段 4｜主体：域内才委托平台内建 / segment 4, delegate the built-in only inside the domain
FC_DL_DintEpochToDt := DINT_TO_DT(nWork);     // 内建还原：纪元秒 → 时刻 / built-in conversion from epoch seconds to an instant
bValid := TRUE;                               // 域内还原可用 / the in-domain instant is usable

// 段 5｜域端点提示（信息级，不置 bError）/ segment 5, domain endpoint hint at info level
IF (nWork = DL_EPOCH_SEC_ZERO) OR (nWork = DL_EPOCH_SEC_MAX) THEN
    eErr := 16#0001_040E;                     // 信息级：输入恰为域端点，多为上游哨兵值 / info level, a domain endpoint, often an upstream sentinel
END_IF
END_FUNCTION

(* ---- FC_DL_DintMsToTime.st ---- *)
(*
    FC_DL_DintMsToTime —— DINT 毫秒到 TIME 防御转换（负值钳零）
    ------------------------------------------------------------------
    分类      : DL_MathData / TimeConv
    前缀      : FC_DL_
    版本      : 1.0.0
    溯源      : IEC 61131-3 标准语义的道莅防御性实现
                （接口语义由 IEC 61131-3 定义，内部委托平台内建 DINT_TO_TIME，
                  外围统一错误码 / 钳位 / 双语文档；clean-room 重写，
                  未复制任何闭源厂商源码，参考实现仅限 MIT/Apache 许可）
    平台      : 纯 IEC 61131-3，CODESYS / TwinCAT / InoProShop 通用
    作者      : 道莅代码库 · PLC编程专家（R17）
    ------------------------------------------------------------------
    功能说明  : 将 DINT 毫秒数防御性转换为 TIME 并作为返回值输出，域内委托平台内建 DINT_TO_TIME；
                负值（TIME 无负语义）钳为 T#0S 并置信息级 16#0001_01F4；
                上溢结构性不可能：DINT 正域上限 2147483647 ms 小于 TIME 域上限 4294967295 ms，
                故本件不设上界饱和分支（该结论已在此声明，后续轮次不得误加上溢假分支）；
                钳位方向：下界钳 0 ms，上界无需要钳；
                纯值类型域无 NaN/±INF 态，故无故障级路径（三个故障槽预留）。
    错误码    : 16#0001_01F4 负毫秒输入（TIME 无负语义），已钳 T#0S——信息级，正常防御
                16#0001_01F5 预留禁用（信息级，不得挪用）
                16#0001_02DC 预留禁用（故障级，不得挪用）
                16#0001_02DD 预留禁用（故障级，不得挪用）
                16#0001_02DE 预留禁用（故障级，不得挪用）
    状态机    : R6 标注 N/A —— 本组件为纯函数无顺序状态机，无 CASE 可写，非法状态不可能出现，故以本节说明替代 ELSE 兜底
    修订记录  : 2026-11-16 v1.0.0 首次入库（R17）
*)
FUNCTION FC_DL_DintMsToTime : TIME
VAR_INPUT
    nMs : DINT; // 毫秒数，有效域 0 ~ 2147483647 ms（负值钳 0） [ms] / milliseconds, valid domain 0 .. 2147483647 ms, negative clamps to 0 [ms]
END_VAR
VAR_OUTPUT
    eErr   : UDINT; // 错误码，0=正常 / error id, 0=ok
    bError : BOOL;  // 是否出错，eErr 非 0 时为 TRUE / error flag, TRUE when eErr is nonzero
    bValid : BOOL;  // 输出是否有效可用 / output valid flag
END_VAR
VAR CONSTANT
    DL_TIME_ZERO : TIME := T#0S; // TIME 零值（负值钳位结果与故障缺省） [ms] / TIME zero value, negative clamp and fault default [ms]
END_VAR

// 段 1｜返回值与错误状态预置 / segment 1, preset return value and error status
FC_DL_DintMsToTime := DL_TIME_ZERO; // 故障缺省返回 T#0S（TIME 无负语义） [ms] / fault default T#0S, TIME has no negative semantics [ms]
eErr   := 0;     // 预置无错误 / preset no error
bError := FALSE; // 预置无故障（本件无故障级路径） / preset no fault, no fault-level path here
bValid := FALSE; // 预置输出无效，通过负值闸后置位 / preset invalid, set TRUE after the negative gate

// 段 2｜负值防御闸（TIME 无负语义） / segment 2, negative guard (TIME has no negative semantics)
IF nMs < 0 THEN
    FC_DL_DintMsToTime := DL_TIME_ZERO; // 负值钳为 T#0S [ms] / clamp the negative value to T#0S [ms]
    eErr := 16#0001_01F4;               // 信息级：负毫秒已钳零，正常防御 / info level: negative milliseconds clamped to zero
    bError := FALSE;                    // 信息级不置故障 / info level never raises fault
    bValid := TRUE;                     // 钳位值本身有效可用 / the clamped value itself is valid
    RETURN;                             // 钳位即出口，不调用内建转换 / clamping is the exit, built-in conversion not called
END_IF

// 段 3｜域内委托转换（末段） / segment 3, in-domain delegated conversion (final)
FC_DL_DintMsToTime := DINT_TO_TIME(nMs); // 域内委托平台内建 DINT_TO_TIME（DINT 正域恒小于 TIME 域，无上溢路径） [ms] / in-domain delegate to built-in DINT_TO_TIME, DINT positive range is always below the TIME range so no overflow path [ms]
eErr   := 0;     // 域内无错误 / in-domain, no error
bError := FALSE; // 信息级不置故障 / info level never raises fault
bValid := TRUE;  // 域内输出有效可用 / in-domain output is valid
END_FUNCTION
